# B&R Automation Studio project DemoCNC
Automation Studio 6.7.0.187; technology packages: mappCockpit 6.7.0, mappMotion 6.7.2, mappView 6.7.0, OpcUaCs 6.0.0

## Configuration Config1

CPU X20CP1684, AutomationRuntime 6.7.6, Build 11.3.0, Vc 6.0.0

### Task classes (Cpu.sw)
```
Cyclic#1 (cycle 2000 us, tolerance 0 us):
  Main <- Cnc.Main.prg
  AxisManual <- Motion.AxisManual.prg
  Handwheel <- Motion.Handwheel.prg
  RingBuffer <- Motion.RingBuffer.prg
  Dispenser <- Heads.Dispenser.prg
  Laser <- Heads.Laser.prg
  OpMode <- Cnc.OpMode.prg
Cyclic#4:
  PrgShare <- Cnc.PrgShare.prg
DataObjects: McAcpSys
NcDataObjects: McDriveLog
Binaries: udbdef, ArSvcReg, FWRules, McProfGen, McAcpSim, mvLoader, McAcpDrv, TCData, iomap, Config_4, asfw, Config_3, Settings, Role, Config_6, Config_2, mCoWebSc, User, UaCsConfig, BRRole, Config_5, Config_1, asnxdb1, arconfig, ashwac, ashwd, sysconf
Libraries: runtime, AsZip, FileIO, McBase, MpBase, McAxGroup, McAcpAx, McAxis, McPathGen, MpAxis, McProgInt, McPureVAx, MpCnc, CoTrace, standard, ArSsl, powerlnk, AsIecCon, UaCoal, sys_lib, astime, UaCoalPrv, AsEPL
```

### Hardware
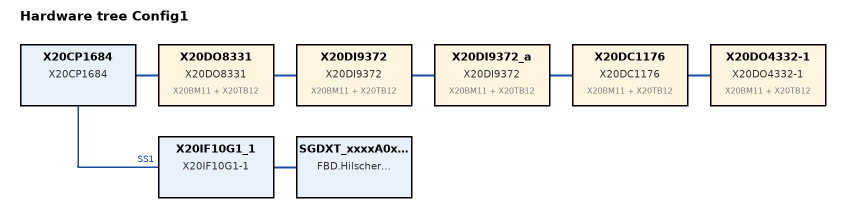
```
SGDXT_xxxxA0x_CoE_Drive_V5_1 : FBD.Hilscher.ECATGenSlaveDTM.SGDXT-xxxxA0x CoE Drive V5.1 v5.1 (OrderNumber=SGDXT-xxxxA0x CoE Drive V5.1)  [ECAT1 -> X20IF10G1_1.IF1]
  DtmId = 5cc0e974-dd08-4d3b-8861-9af8db60d9c1
  ChannelBlocks_556a5014-3061-476e-952f-13eb48db60da  // 2nd_Receive_PDO_mapping_ChA   [OUT, 6 Byte(s)]
  ChannelBlocks_c08b9fef-1a5d-4400-99d8-8c6c7c6492c0  // 2nd_Receive_PDO_mapping_ChB   [OUT, 6 Byte(s)]
  ChannelBlocks_bb719693-a827-4383-9817-184275cbd3ab  // 2nd_Receive_PDO_mapping_ChC   [OUT, 6 Byte(s)]
  ChannelBlocks_bb52f712-f110-4765-9ae9-fe54bf8f2216  // 2nd_Transmit_PDO_mapping_ChA   [IN, 6 Byte(s)]
  ChannelBlocks_06cbf0f9-47c2-45b5-ab43-e0b9d19c4fe2  // 2nd_Transmit_PDO_mapping_ChB   [IN, 6 Byte(s)]
  ChannelBlocks_3a11469b-f58f-4501-9f2d-befe904e9021  // 2nd_Transmit_PDO_mapping_ChC   [IN, 6 Byte(s)]
X20BM11 : X20BM11 v1.1.0.0  [X2X1 -> X20BM11_a.X2X2]
X20BM11_a : X20BM11 v1.1.0.0  [X2X1 -> X20CP1684.IF6]
X20BM11_b : X20BM11 v1.1.0.0  [X2X1 -> X20BM11.X2X2]
X20BM11_c : X20BM11 v1.1.0.0  [X2X1 -> X20BM11_b.X2X2]
X20BM11_d : X20BM11 v1.1.0.0  [X2X1 -> X20BM11_c.X2X2]
X20CP1684 : X20CP1684 v1.9.0.0
  Connector IF2:
    ActivateDevice = 1
    Mode = Manual
    InternetAddress = 192.0.2.10
    SubnetMask = 255.255.255.0
  ConfigurationID = first_Config1
  TimerDeviceType = EPLX2X
  TimerDevice = X20CP1684.IF6
  TaskClassIdleTime = 2000
  Cyclic1Duration = 2000
  Cyclic1Tolerance = 0
  FileDevice1
  FileDeviceName1 = USER
  FileDevicePath1 = USER_PATH
  ActivateWebServer = 1
  ActivateSdm = 1
  Authentication = 0
X20DC1176 : X20DC1176 v1.4.2.0  [SS1 -> X20TB12_c.SS; SL -> X20BM11_c.SL1]
  Supervision = off
  CounterStd01 = 32Bit
  ABRInputs = on
  BrokenWireConfig = off
X20DI9372 : X20DI9372 v1.6.1.0  [SS1 -> X20TB12.SS; SL -> X20BM11.SL1]
  Supervision = off
X20DI9372_a : X20DI9372 v1.6.1.0  [SS1 -> X20TB12_b.SS; SL -> X20BM11_b.SL1]
  Supervision = off
X20DO4332-1 : X20DO4332-1 v1.7.1.0  [SS1 -> X20TB12_d.SS; SL -> X20BM11_d.SL1]
  Supervision = off
X20DO8331 : X20DO8331 v1.2.2.0  [SS1 -> X20TB12_a.SS; SL -> X20BM11_a.SL1]
  Supervision = off
X20IF10G1_1 : X20IF10G1-1 v1.0.2.0  [SS -> X20CP1684.SS1]
  Connector IF1:
    DtmRef = FBDIF.Hilscher.ECATMasterDTM.NETX 100 RE/ECM
    DtmId = 1a6e2b8c-b0d3-41a0-9abf-558976bc5f68
  ConfigFile = X20IF10G1_1.dtm
  ConfigModule = asnxdb1
  CycleTime = 2000
  Synchron = on
X20TB12 : X20TB12 v1.0.0.0
X20TB12_a : X20TB12 v1.0.0.0
X20TB12_b : X20TB12 v1.0.0.0
X20TB12_c : X20TB12 v1.0.0.0
X20TB12_d : X20TB12 v1.0.0.0
```

### BRRole.brrole - X20CP1684/AccessAndSecurity/UserRoleSystem/BRRole.brrole
```
Element BR_Anonymous (Type=BRRole)
Element BR_Engineer (Type=BRRole)
Element BR_Observer (Type=BRRole)
Element BR_SafetyAdmin (Type=BRRole)
Element BR_SecurityAdmin (Type=BRRole)
```

### IoMap.iom - X20CP1684/IoMap.iom
```iecst
VAR_CONFIG
	::gDS402_X.ControlWord AT %QW."SGDXT_xxxxA0x_CoE_Drive_V5_1".2nd_Receive_PDO_mapping_ChA_Control_word;
	::gDS402_X.TargetPosition AT %QD."SGDXT_xxxxA0x_CoE_Drive_V5_1".2nd_Receive_PDO_mapping_ChA_Target_position;
	::gDS402_Y.ControlWord AT %QW."SGDXT_xxxxA0x_CoE_Drive_V5_1".2nd_Receive_PDO_mapping_ChB_Control_word;
	::gDS402_Y.TargetPosition AT %QD."SGDXT_xxxxA0x_CoE_Drive_V5_1".2nd_Receive_PDO_mapping_ChB_Target_position;
	::gDS402_Z.ControlWord AT %QW."SGDXT_xxxxA0x_CoE_Drive_V5_1".2nd_Receive_PDO_mapping_ChC_Control_word;
	::gDS402_Z.TargetPosition AT %QD."SGDXT_xxxxA0x_CoE_Drive_V5_1".2nd_Receive_PDO_mapping_ChC_Target_position;
	::gDS402_X.StatusWord AT %IW."SGDXT_xxxxA0x_CoE_Drive_V5_1".2nd_Transmit_PDO_mapping_ChA_Status_word;
	::gDS402_X.ActualPosition AT %ID."SGDXT_xxxxA0x_CoE_Drive_V5_1".2nd_Transmit_PDO_mapping_ChA_Position_actual_value;
	::gDS402_Y.StatusWord AT %IW."SGDXT_xxxxA0x_CoE_Drive_V5_1".2nd_Transmit_PDO_mapping_ChB_Status_word;
	::gDS402_Y.ActualPosition AT %ID."SGDXT_xxxxA0x_CoE_Drive_V5_1".2nd_Transmit_PDO_mapping_ChB_Position_actual_value;
	::gDS402_Z.StatusWord AT %IW."SGDXT_xxxxA0x_CoE_Drive_V5_1".2nd_Transmit_PDO_mapping_ChC_Status_word;
	::gDS402_Z.ActualPosition AT %ID."SGDXT_xxxxA0x_CoE_Drive_V5_1".2nd_Transmit_PDO_mapping_ChC_Position_actual_value;
	::gDS402_X.DigitalInputs.NegativeLimitSwitch AT %IX."X20DI9372".DigitalInput01;
	::gDS402_X.DigitalInputs.HomingSwitch AT %IX."X20DI9372".DigitalInput02;
	::gDS402_X.DigitalInputs.PositiveLimitSwitch AT %IX."X20DI9372".DigitalInput03;
	::gDS402_Y.DigitalInputs.NegativeLimitSwitch AT %IX."X20DI9372".DigitalInput04;
	::gDS402_Y.DigitalInputs.HomingSwitch AT %IX."X20DI9372".DigitalInput05;
	::gDS402_Y.DigitalInputs.PositiveLimitSwitch AT %IX."X20DI9372".DigitalInput06;
	::gDS402_Z.DigitalInputs.NegativeLimitSwitch AT %IX."X20DI9372".DigitalInput07;
	::gDS402_Z.DigitalInputs.HomingSwitch AT %IX."X20DI9372".DigitalInput08;
	::gDS402_Z.DigitalInputs.PositiveLimitSwitch AT %IX."X20DI9372".DigitalInput09;
	::DO_Dispenser_Start AT %QX."X20DO8331".DigitalOutput01;
	::DO_Laser_Power AT %QX."X20DO8331".DigitalOutput02;
	::PWM_Laser_Duty AT %QW."X20DO4332-1".PwmOutput01;
	::PWM_Laser_Period AT %QW."X20DO4332-1".PwmPeriode;
	::Handwheel:counterValue AT %ID."X20DC1176".Encoder01;
	::Handwheel:counterReset AT %QX."X20DC1176".Encoder01Reset;
	::DI_MPG_AxisX AT %IX."X20DI9372_a".DigitalInput01;
	::DI_MPG_AxisY AT %IX."X20DI9372_a".DigitalInput02;
	::DI_MPG_AxisZ AT %IX."X20DI9372_a".DigitalInput03;
	::DI_MPG_X1 AT %IX."X20DI9372_a".DigitalInput05;
	::DI_MPG_X10 AT %IX."X20DI9372_a".DigitalInput06;
	::DI_MPG_X100 AT %IX."X20DI9372_a".DigitalInput07;
	::DI_MPG_Jog_EMS1 AT %IX."X20DI9372_a".DigitalInput08;
END_VAR
```

- Physical/Config1/X20CP1684/PvMap.vvm: same as Physical/Config1/X20CP1684/Cpu.per
### Config_1.axesgroup - X20CP1684/mappMotion/3AxesCNCXYZ/Config_1.axesgroup
```
Element gCncXYZ (Type=axesgroup)
  Type = PathGenAxesGroup
    PhysicalAxes:
      JointAxes:
        JointAxis[1]:
          Name = QX
          AxisRef = gAxis_X
        JointAxis[2]:
          Name = QY
          AxisRef = gAxis_Y
        JointAxis[3]:
          Name = QZ
          AxisRef = gAxis_Z
    MechanicalSystem:
      MechSysRef = MechSys_3AxCNCXYZ
    AxesGroupFeatures:
      FeatureRef[1] = Feature_Programs
      FeatureRef[2] = Feature_Jogging
      FeatureRef[3] = Feature_MFunctions
      FeatureRef[4] = Feature_HomingOrder
      FeatureRef[5] = Feature_PrgSimAndRestart
```

### Config_2.axis - X20CP1684/mappMotion/3AxesCNCXYZ/Config_2.axis
```
Element gAxis_X (Type=axis)
  BaseType = LinearBounded
    MeasurementResolution = 0.001
    CountDirection = Inverse
  MovementLimits:
    Position:
      LowerLimit = -5
      UpperLimit = 450
    Velocity:
      Velocity = 200
    Acceleration:
      Acceleration = 500.0
    Deceleration:
      Deceleration = 500.0
Element gAxis_Y (Type=axis)
  BaseType = LinearBounded
    MeasurementResolution = 0.001
    CountDirection = Inverse
  MovementLimits:
    Position:
      LowerLimit = -5
      UpperLimit = 430
    Velocity:
      Velocity = 200
    Acceleration:
      Acceleration = 500.0
    Deceleration:
      Deceleration = 500.0
Element gAxis_Z (Type=axis)
  BaseType = LinearBounded
    MeasurementResolution = 0.001
  MovementLimits:
    Position:
      LowerLimit = -5
      UpperLimit = 145
    Velocity:
      Velocity = 200
    Acceleration:
      Acceleration = 500.0
    Deceleration:
      Deceleration = 500.0
```

### Config_3.mechanicalsystem - X20CP1684/mappMotion/3AxesCNCXYZ/Config_3.mechanicalsystem
```
Element MechSys_3AxCNCXYZ (Type=mechanicalsystem)
  Type = 3AxesCNC
    Subtype:
      JointAxesPositionLimits:
        JointAxis[1]
        JointAxis[2]
        JointAxis[3]
```

### Config_4.axesgroupfeature - X20CP1684/mappMotion/3AxesCNCXYZ/Config_4.axesgroupfeature
```
Element Feature_Programs (Type=axesgroupfeature)
  Type = Program
    ModalDataBehaviour = UseAxesGroupSettings
    InitialSettings:
      InterpolationTypes = LinearRapid
      PositionCoordinates = Absolute
      CircleCoordinates = Relative
      JACS_ACSProgramming = JACS
      ContourConnection = Inactive
      AccuracyHoldDelays = None
      ProgrammingUnits = UseAxesGroupSettings
      Feedrates:
        FeedPath = Standard
        FeedCharacteristic = StandardCharacteristic
        FeedType = Feedrate
        FeedReduction = Inactive
        FeedrateValue = 0.0
        InverseFeedrateValue = 0.0
        FeedratePerRevValue = 0.0
    ProgramElements:
      PVs:
        PV[1]:
          PvName = ::C_LaserPower
          Advanced:
            Alias = LaserPower
            Synchronization = Path
        PV[2]:
          PvName = ::C_TP1_1
          Advanced:
            Alias = TP1_1
        PV[3]:
          PvName = ::C_TP1_2
          Advanced:
            Alias = TP1_2
        PV[4]:
          PvName = ::C_TP1_3
          Advanced:
            Alias = TP1_3
        PV[5]:
          PvName = ::C_TP2_1
          Advanced:
            Alias = TP2_1
        PV[6]:
          PvName = ::C_TP2_2
          Advanced:
            Alias = TP2_2
        PV[7]:
          PvName = ::C_TP2_3
          Advanced:
            Alias = TP2_3
        PV[8]:
          PvName = ::C_TP3_1
          Advanced:
            Alias = TP3_1
        PV[9]:
          PvName = ::C_TP3_2
          Advanced:
            Alias = TP3_2
        PV[10]:
          PvName = ::C_TP3_3
          Advanced:
            Alias = TP3_3
        PV[11]:
          PvName = ::C_TP4_1
          Advanced:
            Alias = TP4_1
        PV[12]:
          PvName = ::C_TP4_2
          Advanced:
            Alias = TP4_2
        PV[13]:
          PvName = ::C_TP4_3
          Advanced:
            Alias = TP4_3
    DefaultLanguage = BRGCode
    Location = Default
      FileDevice = CNC_PrgDir
Element Feature_Jogging (Type=axesgroupfeature)
  Type = Jogging
```

### Config_5.purevaxcfg - X20CP1684/mappMotion/3AxesCNCXYZ/Config_5.purevaxcfg
```
Element PureVAxCfg_X (Type=purevaxcfg)
  PureVAxis:
    AxisReference = gAxis_X
    Homing:
      Mode = SwitchGate
        SwitchEdge = Negative
        StartDirection = Negative
    GeneralPurposeAxisInterface = DS402CSP
      MechanicalElements:
        RotaryToLinearTransformation:
          ReferenceDistance = 10
      EncoderSettings:
        IncrementsPerRevolution = 1048576
      PositionActualValue:
        Source = Variable
          PVMapping = ::gDS402_X.ActualPosition
      DigitalInputs:
        HomingSwitch:
          Source = InputPV
            PVmapping = ::gDS402_X.DigitalInputs.HomingSwitch
        PositiveLimitSwitch:
          Source = InputPV
            PVmapping = ::gDS402_X.DigitalInputs.PositiveLimitSwitch
          Level = Low
        NegativeLimitSwitch:
          Source = InputPV
            PVmapping = ::gDS402_X.DigitalInputs.NegativeLimitSwitch
          Level = Low
      StatusInputs:
        StatusWord:
          Source = InputPV
            PVmapping = ::gDS402_X.StatusWord
        ErrorCode:
          Source = InputPV
            PVmapping = ::gDS402_X.ErrorCode
      ControlOutputs:
        ControlWord:
          Destination:
            PVMapping = ::gDS402_X.ControlWord
        TargetPosition:
          Destination:
            PVmapping = ::gDS402_X.TargetPosition
Element PureVAxCfg_Y (Type=purevaxcfg)
  PureVAxis:
    AxisReference = gAxis_Y
    Homing:
      Mode = SwitchGate
        Position = 0
        SwitchEdge = Negative
        StartDirection = Negative
    GeneralPurposeAxisInterface = DS402CSP
      MechanicalElements:
        RotaryToLinearTransformation:
          ReferenceDistance = 10
      EncoderSettings:
        IncrementsPerRevolution = 1048576
      PositionActualValue:
        Source = Variable
          PVMapping = ::gDS402_Y.ActualPosition
      DigitalInputs:
        HomingSwitch:
          Source = InputPV
            PVmapping = ::gDS402_Y.DigitalInputs.HomingSwitch
        PositiveLimitSwitch:
          Source = InputPV
            PVmapping = ::gDS402_Y.DigitalInputs.PositiveLimitSwitch
          Level = Low
        NegativeLimitSwitch:
          Source = InputPV
            PVmapping = ::gDS402_Y.DigitalInputs.NegativeLimitSwitch
          Level = Low
      StatusInputs:
        StatusWord:
          Source = InputPV
            PVmapping = ::gDS402_Y.StatusWord
        ErrorCode:
          Source = InputPV
            PVmapping = ::gDS402_Y.ErrorCode
      ControlOutputs:
        ControlWord:
          Destination:
            PVMapping = ::gDS402_Y.ControlWord
        TargetPosition:
          Destination:
            PVmapping = ::gDS402_Y.TargetPosition
Element PureVAxCfg_Z (Type=purevaxcfg)
  PureVAxis:
    AxisReference = gAxis_Z
    Homing:
      Mode = SwitchGate
        SwitchEdge = Negative
        StartDirection = Negative
    GeneralPurposeAxisInterface = DS402CSP
      MechanicalElements:
        RotaryToLinearTransformation:
          ReferenceDistance = 10
      EncoderSettings:
        IncrementsPerRevolution = 1048576
      PositionActualValue:
        Source = Variable
          PVMapping = ::gDS402_Z.ActualPosition
      DigitalInputs:
        HomingSwitch:
          Source = InputPV
            PVmapping = ::gDS402_Z.DigitalInputs.HomingSwitch
        PositiveLimitSwitch:
          Source = InputPV
            PVmapping = ::gDS402_Z.DigitalInputs.PositiveLimitSwitch
          Level = Low
        NegativeLimitSwitch:
          Source = InputPV
            PVmapping = ::gDS402_Z.DigitalInputs.NegativeLimitSwitch
          Level = Low
      StatusInputs:
        StatusWord:
          Source = InputPV
            PVmapping = ::gDS402_Z.StatusWord
        ErrorCode:
          Source = InputPV
            PVmapping = ::gDS402_Z.ErrorCode
      ControlOutputs:
        ControlWord:
          Destination:
            PVMapping = ::gDS402_Z.ControlWord
        TargetPosition:
          Destination:
            PVmapping = ::gDS402_Z.TargetPosition
```

### Config_6.axesgroupfeature - X20CP1684/mappMotion/3AxesCNCXYZ/Config_6.axesgroupfeature
```
Element Feature_MFunctions (Type=axesgroupfeature)
  Type = MFunctions
    MFunction[1]:
      IndexType = Range
        IndexFrom = 40
        IndexTo = 49
      Blocking = Disabled
    MFunction[2]:
      IndexType = Range
        IndexFrom = 50
        IndexTo = 59
    MFunction[3]:
      IndexType = Range
        IndexFrom = 60
        IndexTo = 69
      Blocking = Disabled
```

### Config_7.axesgroupfeature - X20CP1684/mappMotion/3AxesCNCXYZ/Config_7.axesgroupfeature
```
Element Feature_HomingOrder (Type=axesgroupfeature)
  Type = HomingOrder
    TogetherGroup[1]:
      AxisRef[1] = gAxis_Z
    TogetherGroup[2]:
      AxisRef[1] = gAxis_X
      AxisRef[2] = gAxis_Y
```

### Config_8.axesgroupfeature - X20CP1684/mappMotion/3AxesCNCXYZ/Config_8.axesgroupfeature
```
Element Feature_PrgSimAndRestart (Type=axesgroupfeature)
  Type = SimulationRestart
    ConditionalStop = NotUsed
    AdvancedParameters = NotUsed
```

## Logical view

Binary libraries used (declarations not repeated): operator, runtime, AsIecCon, astime, AsZip, FileIO, McBase 6.7.2, MpBase 6.5.0, McAxGroup 6.7.2, McAcpAx 6.7.2, McAxis 6.7.2, McPathGen 6.7.2, MpAxis 6.7.2, McProgInt 6.7.2, McPureVAx 6.7.2, MpCnc 6.7.2, CoTrace 6.7.0, standard

### Global.typ - Global data types
```iecst
TYPE
	Equip_Type : 	STRUCT
		Input : EquipInput_Type;
		Output : EquipOutput_Type;
	END_STRUCT;
	EquipInput_Type : 	STRUCT
		Command : EquipInputCommand_Type;
		CncCommand : E_CNC_ACTION;
		Parameter : EquipInputParameter_Type;
	END_STRUCT;
	EquipOutput_Type : 	STRUCT
		State : EquipOutputState_Type;
		Status : EquipOutputStatus_Type;
	END_STRUCT;
	EquipInputCommand_Type : 	STRUCT
		ManualMove : BOOL; (*move to Parameter.ManualPositon (Z retracts to 0 first) - manual mode, homed*)
		AlarmClearAll : BOOL;
		ManualMode : BOOL; (*TRUE = manual mode (jog, position move, manual discharge). Ignored while the CNC is busy*)
	END_STRUCT;
	EquipInputParameter_Type : 	STRUCT
		sProgramName : STRING[80];
		DryRun : BOOL;
		SystemSpeed : REAL;
		Feedrate : REAL;
		ManualSlowMove : BOOL;
		ManualPositon : ARRAY[0..2]OF REAL;
		sBlock : STRING[260]; (*single NC block for E_ACT_MOVE_BLOCK (MDI), e.g. 'G90 G01 X10 Y20 F1000'*)
		sInitProgram : STRING[80]; (*init program run before every program START (not MDI) as an init subroutine of the program (MoveProgramOptions.InitProgram), e.g. a G92 or a move to a teach position. Empty = none*)
	END_STRUCT;
	EquipOutputState_Type : 	STRUCT
		Initialized : BOOL;
		Stop : BOOL;
		Move : BOOL;
		Complete : BOOL;
	END_STRUCT;
	EquipOutputStatus_Type : 	STRUCT
		CurrentAction : E_CNC_ACTION;
		Mode : BOOL;
		ManualMove : BOOL;
		MoveComplete : BOOL;
		WorkPanelName : STRING[255];
		PowerOn : BOOL; (*CNC axes powered*)
		IsHomed : BOOL; (*CNC axes homed - FALSE after every power-up until HOME / INIT*)
		ProgramActive : BOOL; (*CNC program executing (also while interrupted)*)
		ProgramInterrupted : BOOL; (*CNC program interrupted by HALT*)
		Error : BOOL; (*MpCnc3Axis error*)
		StatusID : DINT; (*MpCnc3Axis StatusID*)
		Rejected : E_CNC_ACTION; (*last mailbox command discarded because its preconditions were not met, IDLE after an accepted command*)
		EmergencyStop : BOOL; (*E-stop latched - release the button, then RESET*)
	END_STRUCT;
	E_CNC_ACTION :
		(
		E_ACT_IDLE := 0,
		E_ACT_INIT := 1,
		E_ACT_START := 2,
		E_ACT_HALT := 3,
		E_ACT_STOP := 4,
		E_ACT_RESET := 5,
		E_ACT_CONTINUE := 6,
		E_ACT_LOADPROGRAM := 7,
		E_ACT_HOME := 8,
		E_ACT_ABORT := 10, (*leave the running command without an action (Main), refused while idle*)
		E_ACT_POWER_OFF := 13, (*servo off*)
		E_ACT_MOVE_BLOCK := 14, (*execute Parameter.sBlock (MDI)*)
		E_ACT_START_AT_LINE := 15, (*START from the file line gCncRun.Input.StartLine*)
		E_ACT_MEASURE_Z := 16 (*Z reference measurement with the touch sensor (gZRef) - manual mode, homed*)
		);
END_TYPE

(*Dispenser*)

TYPE
	Dispenser_Type : 	STRUCT
		Input : DispenserInput_Type;
		Output : DispenserOutput_Type;
	END_STRUCT;
	DispenserInput_Type : 	STRUCT
		Command : DispenserInputCommand_Type;
		Parameter : DispenserInputParameter_Type;
	END_STRUCT;
	DispenserOutput_Type : 	STRUCT
		State : DispenserOutputState_Type;
	END_STRUCT;
	DispenserInputCommand_Type : 	STRUCT
		Discharge : BOOL; (*auto : M41 on / M42 off, driven by Main*)
		Manual : BOOL; (*manual on/off*)
	END_STRUCT;
	DispenserInputParameter_Type : 	STRUCT
		DischargeDelay : BOOL; (*M44 on / M45 off - flag for the program, no output function on this machine*)
	END_STRUCT;
	DispenserOutputState_Type : 	STRUCT
		Discharge : BOOL; (*TRUE while the dispenser discharges (DO_Dispenser_Start)*)
	END_STRUCT;
END_TYPE

(*Laser*)

TYPE
	Laser_Type : 	STRUCT
		Input : LaserInput_Type;
		Output : LaserOutput_Type;
	END_STRUCT;
	LaserInput_Type : 	STRUCT
		Command : LaserInputCommand_Type;
		Parameter : LaserInputParameter_Type;
	END_STRUCT;
	LaserOutput_Type : 	STRUCT
		State : LaserOutputState_Type;
	END_STRUCT;
	LaserInputCommand_Type : 	STRUCT
		Emission : BOOL; (*auto : M61 on / M62 off, driven by Main*)
		Manual : BOOL; (*manual on/off*)
	END_STRUCT;
	LaserInputParameter_Type : 	STRUCT (*written by the HMI (gLaser is not RETAIN, the Laser Init sets the start values)*)
		Power : REAL; (*auto power [%] while the program sets no LaserPower (C_LaserPower < 0)*)
		ManualPower : REAL; (*manual test power [%]*)
		DutyMin : REAL; (*PWM duty for a power just above 0 % [%] - lasing threshold of the driver*)
		DutyMax : REAL; (*PWM duty for 100 % power [%]*)
		PwmPeriod : UINT; (*PWM period [us], 1000..65535 (1000 = 1 kHz, the X20DO4332-1 maximum)*)
		SpeedScale : BOOL; (*corner compensation : power x actual / programmed path velocity*)
		MinSpeedRatio : REAL; (*lower limit of that velocity ratio [%]*)
	END_STRUCT;
	LaserOutputState_Type : 	STRUCT
		Emission : BOOL; (*TRUE while the laser emits (DO_Laser_On : on and power > 0)*)
		Power : REAL; (*power output now [%], after corner compensation, 0 while off*)
		Duty : REAL; (*PWM duty output now [%]*)
	END_STRUCT;
END_TYPE

(*Axis*)

TYPE
	AXIS_COMMAND :
		(
		Axis_IDLE := 0,
		Axis_MOVE_ABSOLUTE := 1,
		Axis_STOP := 2,
		Axis_HALT := 3,
		Axis_JOG_NEGATIVE := 4,
		Axis_JOG_POSITIVE := 5,
		Axis_RESET := 6,
		Axis_MOVE_ADDITIVE := 7,
		Axis_HOME := 8,
		Axis_POWER := 9,
		Axis_MOVE_VELOCITY := 10
		);
	AxesInterface_Type : 	STRUCT
		Input : AxisInput_Type;
		Output : AxisOutput_Type;
	END_STRUCT;
	AxisInput_Type : 	STRUCT
		Parameter : AxisParameter_Type;
		Command : AxisCommand_Type;
	END_STRUCT;
	AxisOutput_Type : 	STRUCT
		State : AxisState_Type;
	END_STRUCT;
	AxisCommand_Type : 	STRUCT
		JogNegative : BOOL;
		JogPositive : BOOL;
		Reset : BOOL;
		Command : AXIS_COMMAND;
	END_STRUCT;
	AxisParameter_Type : 	STRUCT
		Speed : REAL;
		Position : REAL;
		Distance : REAL;
		JogSpeed : REAL;
		SoftwareLimitsPos : DINT;
		SoftwareLimitsNeg : DINT;
		Power : BOOL; (*target of Axis_POWER : TRUE = on, FALSE = off*)
	END_STRUCT;
	AxisState_Type : 	STRUCT
		Enable : BOOL;
		Home : BOOL;
		JogNegative : BOOL;
		JogPositive : BOOL;
		Error : BOOL;
		ErrorID : UDINT;
		Status : SINT; (*0: Not Init , 1 : Idle or OK , 2 : Run, 3 : Error *)
		Command : AXIS_COMMAND;
		Position : LREAL;
		Speed : LREAL;
	END_STRUCT;
END_TYPE

(*Drive diagnosis - read-only copies for the HMI, not RETAIN (gAxis is RETAIN and keeps its structure). Written by AxisManual*)

TYPE
	DriveDiag_Type : 	STRUCT
		Valid : BOOL; (*the values below are up to date (MC_ReadAxisInfo.Valid) - FALSE = do not judge them*)
		CommReady : BOOL; (*drive has a network connection (MC_ReadAxisInfo.CommunicationReady) - follows the 'Module ok' status input of the axis config (Config_5), not used yet*)
		ReadyForPowerOn : BOOL; (*drive can be switched on (MC_ReadAxisInfo.ReadyForPowerOn)*)
		Warning : BOOL; (*a warning is active on the drive (MC_ReadAxisInfo.AxisWarning, DS402 status word bit 7)*)
		WarningAlarm : BOOL; (*warning-level alarm for the HMI (alarms.json exType 1) : Warning while Valid and CommReady for 0.5 s, held 2 s after it clears (one alarm per event, no flicker). Display only - the PLC does not react to it*)
	END_STRUCT;
END_TYPE

(*Position move result*)

TYPE
	ManualMoveResult_Type : 	STRUCT (*result of gEquipment.Input.Command.ManualMove, written by AxisManual - its own non-RETAIN global so the RETAIN gEquipment keeps its layout*)
		Result : USINT; (*result of request number Count : 0 none since power-up, 1 running, 2 arrived (every step of the sequence done), 3 refused (dropped, nothing moved), 4 ended before the target (Reason)*)
		Reason : USINT; (*why refused / ended, 0 none : 1 E-stop, 2 auto mode, 3 handwheel selected, 4 CNC command running, 5 axes moving, 6 not homed, 7 servo off, 8 axis error, 9 axis HALT / STOP, 10 an axis move of the sequence was aborted or failed (the sequence went on)*)
		Count : UINT; (*+1 for every ManualMove request the PLC takes (accepted or refused) : a new result also when it equals the last one*)
	END_STRUCT;
END_TYPE

(*Z reference measurement - touch sensor DI_ZRef_Sensor (not wired yet), cycle in Main Action_ZRef.st (CncCommand E_ACT_MEASURE_Z)*)

TYPE
	ZRef_Type : 	STRUCT
		Input : ZRefInput_Type;
		Output : ZRefOutput_Type;
	END_STRUCT;
	ZRefInput_Type : 	STRUCT (*written by the HMI, kept over power off (gZRef is RETAIN) - machine coordinates [mm], Z+ down (0 = top). All 0 = not set : the command is refused*)
		SensorX : LREAL; (*X of the sensor*)
		SensorY : LREAL; (*Y of the sensor*)
		StartZ : LREAL; (*Z above the sensor where the slow search starts*)
		MaxZ : LREAL; (*deepest Z of the search : no signal down to here = failed (at most 50 mm below StartZ)*)
		SafeZ : LREAL; (*Z of the moves to and from the sensor (not below StartZ), usually 0*)
		ProbeVel : REAL; (*search velocity [mm/s], 0 = 2, at most 10. The result is read once per cycle : error up to about ProbeVel x 2 cycles (2 ms) + the input filter*)
		Head : USINT; (*head being measured (HMI head number), copied to Output.Head with the result*)
	END_STRUCT;
	ZRefOutput_Type : 	STRUCT
		ParamOk : BOOL; (*Input valid : SafeZ <= StartZ < MaxZ, search <= 50 mm, all inside the software limits, ProbeVel <= 10*)
		Sensor : BOOL; (*DI_ZRef_Sensor now*)
		Busy : BOOL; (*measurement running*)
		Step : USINT; (*diagnosis: 10 Z to SafeZ, 20 X / Y to the sensor, 30 Z to StartZ, 40 search, 50 braking, 60 Z back to SafeZ*)
		Done : BOOL; (*MeasuredZ is the result of the last measurement (cleared when the next one starts)*)
		MeasuredZ : LREAL; (*Z at the sensor signal [mm, machine]*)
		Head : USINT; (*head of MeasuredZ*)
		ErrorId : USINT; (*last measurement: 0 none, 1 Input not valid, 2 sensor already on at StartZ, 3 no signal down to MaxZ, 4 axis move failed or aborted (jog, axis error), 5 left (STOP, ABORT, E-stop, handwheel), 6 a move did not finish in time*)
	END_STRUCT;
END_TYPE

(*Work offsets G54..G57 - program origin in machine coordinates, set as the standard frame SCS1 before a program / MDI run (Main Action_WorkOffset.st)*)

TYPE
	WorkOffset_Type : 	STRUCT
		Input : WorkOffsetInput_Type;
		Output : WorkOffsetOutput_Type;
	END_STRUCT;
	WorkOffsetInput_Type : 	STRUCT
		Command : WorkOffsetInputCommand_Type;
		Parameter : WorkOffsetInputParameter_Type;
	END_STRUCT;
	WorkOffsetInputCommand_Type : 	STRUCT
		Apply : BOOL; (*pulse: take Parameter over (table and Active), cleared by the PLC - refused while a command / program runs*)
	END_STRUCT;
	WorkOffsetInputParameter_Type : 	STRUCT
		Offset : ARRAY[0..3]OF WorkOffsetXYZ_Type; (*0 = G54 .. 3 = G57 : machine position of the program origin [mm]*)
		Active : USINT; (*0..3 = G54..G57 : offset used by every program and MDI run*)
	END_STRUCT;
	WorkOffsetXYZ_Type : 	STRUCT
		X : LREAL;
		Y : LREAL;
		Z : LREAL;
	END_STRUCT;
	WorkOffsetOutput_Type : 	STRUCT
		Offset : ARRAY[0..3]OF WorkOffsetXYZ_Type; (*table in effect (taken over by Apply, kept over power off)*)
		Active : USINT; (*offset in effect, 0 = G54*)
		InUse : BOOL; (*the frame is set before every run : the active offset or the frame set last is not 0*)
		Rejected : BOOL; (*the last Apply was refused : CNC busy, Active > 3 or a value out of range (10000 mm)*)
		Error : BOOL; (*setting the frame failed - that run was not started*)
		ErrorID : DINT; (*ErrorID of MC_BR_SetStandardFrame, 0 = none*)
	END_STRUCT;
END_TYPE

(*Head (tool) offsets - offset of the mounted head from the reference head tip, set as the standard frame SCS2 before a program / MDI run (Main Action_HeadOffset.st)*)

TYPE
	HeadOffset_Type : 	STRUCT
		Input : HeadOffsetInput_Type;
		Output : HeadOffsetOutput_Type;
	END_STRUCT;
	HeadOffsetInput_Type : 	STRUCT
		Command : HeadOffsetInputCommand_Type;
		Parameter : HeadOffsetInputParameter_Type;
	END_STRUCT;
	HeadOffsetInputCommand_Type : 	STRUCT
		Apply : BOOL; (*pulse: take Parameter over (table and ActiveHead), cleared by the PLC - refused while a command / program runs*)
	END_STRUCT;
	HeadOffsetInputParameter_Type : 	STRUCT
		Offset : ARRAY[1..4]OF HeadOffsetXYZ_Type; (*head 1..4 (HMI head table H1..H4 = plugin PlcId : 1 dispenser, 2 laser) : from the reference head tip (the point the axis positions refer to) to the working point of that head [mm], machine directions (Z+ down)*)
		ActiveHead : USINT; (*mounted head 1..4 whose offset every program and MDI run uses, 0 = none (no offset)*)
	END_STRUCT;
	HeadOffsetXYZ_Type : 	STRUCT
		X : LREAL;
		Y : LREAL;
		Z : LREAL;
	END_STRUCT;
	HeadOffsetOutput_Type : 	STRUCT
		Offset : ARRAY[1..4]OF HeadOffsetXYZ_Type; (*table in effect (taken over by Apply, kept over power off)*)
		ActiveHead : USINT; (*head in effect, 0 = none*)
		InUse : BOOL; (*the frame is set before every run : the active head's offset or the frame set last is not 0*)
		Rejected : BOOL; (*the last Apply was refused : CNC busy, ActiveHead > 4 or a value out of range (1000 mm)*)
		Error : BOOL; (*setting the frame failed - that run was not started*)
		ErrorID : DINT; (*ErrorID of MC_BR_SetStandardFrame, 0 = none*)
	END_STRUCT;
END_TYPE

(*CNC program run options from the HMI (gCncRun, not RETAIN : everything is off after a power-up)*)

TYPE
	CncRun_Type : 	STRUCT
		Input : CncRunInput_Type;
		Output : CncRunOutput_Type;
	END_STRUCT;
	CncRunInput_Type : 	STRUCT
		SingleStep : BOOL; (*TRUE = single step : the program stops after every block, CONTINUE runs the next one (MpCnc3Axis.SingleStep). Not used for MDI*)
		OptionalStop : BOOL; (*TRUE = the program stops at M01, CONTINUE goes on (MC_BR_OptionalStop)*)
		StartLine : UDINT; (*E_ACT_START_AT_LINE : line of the program file to start at, 1 = first line (as C_CurrentLine). Write it before CncCommand 15*)
		ReposVelocityFactor : REAL; (*E_ACT_START_AT_LINE : AxisVelocityFactor of the automatic repositioning to the start point (mcPRGRP_SINGLE_AXIS_AUTOMATIC), Main Init sets 0.1*)
	END_STRUCT;
	CncRunOutput_Type : 	STRUCT
		SingleStepActive : BOOL; (*single step mode active (MpCnc3Axis.SingleStepActive)*)
		OptionalStopActive : BOOL; (*the program stands at M01 (MC_BR_OptionalStop.Interrupting) - CONTINUE goes on*)
		OptionalStopErrorId : DINT; (*ErrorID of MC_BR_OptionalStop, 0 = none - switch OptionalStop off and on again to retry*)
		InterruptStatus : McPrgInfoInterruptEnum; (*why the program is interrupted (MpCnc3Axis Info.Program.InterruptStatus) - for commissioning*)
		ProgramPhase : McPrgPhaseEnum; (*MpCnc3Axis Info.Program.ProgramPhase : start at line = simulation up to the line, repositioning, waiting for CONTINUE, real run*)
	END_STRUCT;
END_TYPE
```

### Global.var - Global variables
```iecst
(*Drive adapter - motor / drive specific.
  On a motor or drive change only this block, IoMap.iom, the mappMotion axis configs and the DTM change.
  Program logic uses only the mapp axis references gAxis_X/Y/Z and the axes group gCncXYZ.*)
VAR
	gDS402_X : McPureVAxDS402CspAdapterPvType;
	gDS402_Y : McPureVAxDS402CspAdapterPvType;
	gDS402_Z : McPureVAxDS402CspAdapterPvType;
END_VAR
VAR RETAIN
	gEquipment : Equip_Type;
	gAxis : ARRAY[0..2] OF AxesInterface_Type;
END_VAR
VAR
	gDispenser : Dispenser_Type;
	gLaser : Laser_Type;
END_VAR
(*Axis index of gAxis, gDriveDiag and the per-axis FB arrays*)
VAR CONSTANT
	AX_X : USINT := 0;
	AX_Y : USINT := 1;
	AX_Z : USINT := 2;
	AX_LAST : USINT := 2; (*highest axis index : FOR i := 0 TO AX_LAST*)
END_VAR
(*Drive diagnosis for the HMI - read only (AxisManual overwrites it every cycle), not RETAIN, index AX_X/AX_Y/AX_Z as gAxis*)
VAR
	gDriveDiag : ARRAY[0..2] OF DriveDiag_Type;
END_VAR
(*HMI jog heartbeat - not RETAIN*)
VAR
	gJogAlive : UINT := 0; (*the HMI changes it every 0.1 s while it jogs; AxisManual stops the jog when it stands still for 0.5 s*)
END_VAR
(*Position move result for the HMI - not RETAIN (gEquipment is RETAIN and keeps its layout)*)
VAR
	gManualMoveResult : ManualMoveResult_Type; (*result of the last Input.Command.ManualMove request, written by AxisManual*)
END_VAR
(*Heads - one head on the machine (HMI plugin structure). Head number = PlcId of the HMI head plugin*)
VAR CONSTANT
	HEAD_DISPENSER : USINT := 1; (*dispenser : M41 / M42 discharge on / off, M44 / M45 discharge delay flag, Dispenser task*)
	HEAD_LASER : USINT := 2; (*PWM laser : M61 / M62 emission on / off, Laser task*)
END_VAR
(*Heads this PLC program has - not RETAIN, read by the HMI*)
VAR
	gHeadSupport : UDINT := 0; (*bit n = head n (HEAD_ constants) has its M functions and outputs here. Fixed, set by Main every cycle. The HMI does not offer a head without its bit*)
END_VAR
(*Active head - written by the HMI, not RETAIN. Not in gEquipment : a new field would change the RETAIN structure*)
VAR
	gActiveHead : USINT := 0; (*head selected on the HMI (HEAD_ constant, the plugin PlcId). Only its M functions and manual on are taken : an M function of another head stops the program, a manual on of another head is dropped (Main act_HeadCheck). 0 = not known yet (PLC restart until the HMI writes it) : no check*)
	gHeadRefused : USINT := 0; (*head whose M function or manual on was refused last because it is not gActiveHead (HEAD_ constants), 0 = none. Cleared when the next run starts or by RESET*)
END_VAR
(*CNC program run options from the HMI (single step, M01 stop, start at line) - not RETAIN : off after every power-up*)
VAR
	gCncRun : CncRun_Type;
END_VAR
(*Setting Variable*)
VAR RETAIN
	SlowMoveVelocity : DINT := 10;
	SlowMoveLength : DINT := 100;
END_VAR
(*Monitor*)
VAR
	C_CurrentLine : DINT := 0; (*line of the running CNC program, from MpCnc3Axis ProgramMonitor*)
	C_OverallRuntime : LREAL := 0.0; (*execution time of the running CNC program [s], from MpCnc3Axis ProgramMonitor - counts from the start (file load included) and holds after the end*)
	C_MovementRuntime : LREAL := 0.0; (*movement time of the running CNC program [s], from MpCnc3Axis ProgramMonitor - file load not included*)
	Torque_X : REAL := 0.0;
	Torque_Y : REAL := 0.0;
	Torque_Z : REAL := 0.0;
END_VAR
(*CNC program variables - written by the program through an alias of the axes group program feature (Config_4, path synchronous)*)
VAR
	C_LaserPower : REAL := -1.0; (*LaserPower = <%> in the program; < 0 = not set (gLaser.Input.Parameter.Power), reset at program end*)
END_VAR
(*Teach positions 1..4 [mm, machine coordinates] - read by CNC programs as TP1_1 .. TP4_3 (aliases in Config_4, _1 = X, _2 = Y, _3 = Z : a name
  must not contain X/Y/Z/F after its first letter - an address letter inside an expression
  splits the expression, e.g. 'X=2930-DoubleBeadY=40'), e.g. in the init program
  (Input.Parameter.sInitProgram) 'G00 X=TP1_1 Y=TP1_2' to go there, or 'G92 X=TP4_1 Y=TP4_2' (G92 = absolute zero offset : teach position 4 becomes the program origin). The HMI owns the values (Config\TeachPositions.xml, slot = order
  in Config\Machine.xml) and writes them here whenever they differ*)
VAR RETAIN
	C_TP1_1 : LREAL := 0.0;
	C_TP1_2 : LREAL := 0.0;
	C_TP1_3 : LREAL := 0.0;
	C_TP2_1 : LREAL := 0.0;
	C_TP2_2 : LREAL := 0.0;
	C_TP2_3 : LREAL := 0.0;
	C_TP3_1 : LREAL := 0.0;
	C_TP3_2 : LREAL := 0.0;
	C_TP3_3 : LREAL := 0.0;
	C_TP4_1 : LREAL := 0.0;
	C_TP4_2 : LREAL := 0.0;
	C_TP4_3 : LREAL := 0.0;
END_VAR
(*Z reference measurement (CncCommand E_ACT_MEASURE_Z, Main Action_ZRef.st) - RETAIN on its own (sensor position), gEquipment is
  not changed. The HMI writes Input (sensor position, search range) and reads Output (MeasuredZ, Done, ErrorId)*)
VAR RETAIN
	gZRef : ZRef_Type;
END_VAR
(*Work offsets G54..G57 (Main Action_WorkOffset.st) - RETAIN on its own, gEquipment is not changed. The HMI writes Input.Parameter
  (machine position of the program origin per offset, active offset) and sets Input.Command.Apply while the CNC is idle; the values
  in effect are Output.Offset / Output.Active. All 0 (the default) = program coordinates are machine coordinates*)
VAR RETAIN
	gWorkOffset : WorkOffset_Type;
END_VAR
(*Head (tool) offsets (Main Action_HeadOffset.st) - RETAIN on its own, gEquipment is not changed. The HMI writes Input.Parameter
  (offset per head from the reference head tip, mounted head) and sets Input.Command.Apply while the CNC is idle; the values in
  effect are Output.Offset / Output.ActiveHead. ActiveHead 0 or offset 0 (the default) = no shift*)
VAR RETAIN
	gHeadOffset : HeadOffset_Type;
END_VAR
(*I/O - wired signals only. Axis limit/home switches go straight to gDS402_* in IoMap.iom*)
VAR
	DI_Auto : BOOL := FALSE;
	DI_MPG_AxisX : BOOL := FALSE;
	DI_MPG_AxisY : BOOL := FALSE;
	DI_MPG_AxisZ : BOOL := FALSE;
	DI_MPG_X1 : BOOL := FALSE;
	DI_MPG_X10 : BOOL := FALSE;
	DI_MPG_X100 : BOOL := FALSE;
	DI_MPG_Jog_EMS1 : BOOL := FALSE;
	DI_MPG_Jog_Enable : BOOL := FALSE;
	DO_Dispenser_Start : BOOL := FALSE;
	DO_Laser_Power : BOOL := FALSE; (*X20DO8331 DO02 - on/off laser output, not used by the PWM laser : held FALSE*)
	PWM_Laser_Duty : INT := 0; (*X20DO4332-1 PwmOutput01 : 0..32767 = 0..100 % of the period (power and on/off)*)
	PWM_Laser_Period : UINT := 1000; (*X20DO4332-1 PwmPeriode [us]*)
END_VAR
(*Z reference touch sensor - NOT wired yet : no channel in Hardware.hw / IoMap.iom. Map it in IoMap.iom once the sensor is wired
  (TRUE = touched : an NC sensor needs a NOT where Main reads it). Until then it stays FALSE and a measurement ends at MaxZ (ErrorId 3)*)
VAR
	DI_ZRef_Sensor : BOOL := FALSE;
END_VAR
(*Laser emitting (on and power > 0) - not wired, for the HMI (head lamp, PLC presence)*)
VAR
	DO_Laser_On : BOOL := FALSE;
END_VAR
```


### Package Logical/Cnc - CNC sequence, operating mode, program folder

### Program Logical/Cnc/Main (IEC) - CNC sequencer (MpCnc3Axis)

#### Init.st - Init code
```iecst
PROGRAM _INIT

	gEquipment.Input.CncCommand := E_ACT_IDLE;

	gEquipment.Output.State.Initialized := FALSE;
	gEquipment.Input.Parameter.SystemSpeed := 200; (* [mm/s] position move speed - axis velocity limit is 200 (mappMotion Config_2) *)
	gEquipment.Input.Parameter.Feedrate := 100;

	(* mapp Motion CNC : static references *)
	fbCnc.MpLink := ADR(gCncXYZ);
	fbCnc.Parameters := ADR(CncParameters);
	fbCnc.Enable := TRUE;
	fbCnc.Override := 100.0;
	fbCnc.RapidOverride := 100.0;
	fbCnc.FeedrateOverride := 100.0;

	(* Jog path limits : adjust to machine limits *)
	CncParameters.Jog.PathLimits.Velocity := 1000.0;			(* [mm/s] *)
	CncParameters.Jog.PathLimits.Acceleration := 5000.0;		(* [mm/s^2] *)
	CncParameters.Jog.PathLimits.Deceleration := 5000.0;		(* [mm/s^2] *)

	(* M-Functions : async (AxesGroup M-function feature, ranges 40..49 / 60..69 non-blocking), M50 / M51 blocking (50..59, no function) *)
	fbMFunction[0].MFunction := 41;
	fbMFunction[1].MFunction := 42;
	fbMFunction[2].MFunction := 44;
	fbMFunction[3].MFunction := 45;
	fbMFunction[4].MFunction := 61;
	fbMFunction[5].MFunction := 62;
	fbMFunction[6].MFunction := 50;
	fbMFunction[7].MFunction := 51;
	FOR i := 0 TO 7 DO
		fbMFunction[i].AxesGroup := ADR(gCncXYZ);
		fbMFunction[i].Enable := TRUE;
	END_FOR
	(* M52..M59 : no function here too, act_MSpare lets the path go on (blocking codes of the range would wait for ever) *)
	FOR i := 0 TO 7 DO
		fbMFunctionSpare[i].MFunction := USINT_TO_UDINT(52 + i);
		fbMFunctionSpare[i].AxesGroup := ADR(gCncXYZ);
		fbMFunctionSpare[i].Enable := TRUE;
	END_FOR

	(* Optional stop (M01) : enabled from the HMI (gCncRun.Input.OptionalStop) in Cyclic *)
	fbOptStop.AxesGroup := ADR(gCncXYZ);
	(* Start at line : velocity factor of the automatic single-axis repositioning to the start point - slow on purpose, check on site *)
	gCncRun.Input.ReposVelocityFactor := 0.1;

	(* Z reference measurement (act_MeasureZ) : own single-axis FBs. gZRef.Input (RETAIN) is kept *)
	fbZrMove[0].Axis := ADR(gAxis_X);
	fbZrMove[1].Axis := ADR(gAxis_Y);
	fbZrMove[2].Axis := ADR(gAxis_Z);
	fbZrHalt[0].Axis := ADR(gAxis_X);
	fbZrHalt[1].Axis := ADR(gAxis_Y);
	fbZrHalt[2].Axis := ADR(gAxis_Z);
	FOR i := 0 TO 2 DO
		fbZrMove[i].Acceleration := C_ZREF_ACC;
		fbZrMove[i].Deceleration := C_ZREF_ACC;
		fbZrHalt[i].Deceleration := C_ZREF_ACC;
	END_FOR
	gZRef.Output.Busy := FALSE;
	gZRef.Output.Step := 0;

	(* Work offsets G54..G57 : the active one is set as standard frame SCS1 before a run (act_WorkOffset).
	   The table (gWorkOffset, RETAIN) is kept; the axes group starts with frame 0, so woSet starts at 0 *)
	fbWorkFrame.AxesGroup := ADR(gCncXYZ);
	fbWorkFrame.CoordSystem := mcSCS1;
	fbWorkFrame.ExecutionMode := mcEM_IMMEDIATELY;
	gWorkOffset.Input.Command.Apply := FALSE;
	gWorkOffset.Output.Rejected := FALSE;
	gWorkOffset.Output.Error := FALSE;
	gWorkOffset.Output.ErrorID := 0;

	(* Head (tool) offsets : minus the mounted head's offset is set as standard frame SCS2 before a run (act_HeadOffset).
	   The table (gHeadOffset, RETAIN) is kept; the axes group starts with frame 0, so hoSet starts at 0 *)
	fbHeadFrame.AxesGroup := ADR(gCncXYZ);
	fbHeadFrame.CoordSystem := mcSCS2;
	fbHeadFrame.ExecutionMode := mcEM_IMMEDIATELY;
	gHeadOffset.Input.Command.Apply := FALSE;
	gHeadOffset.Output.Rejected := FALSE;
	gHeadOffset.Output.Error := FALSE;
	gHeadOffset.Output.ErrorID := 0;

	(* Axis reset FBs *)
	fbAxisReset[0].Axis := ADR(gAxis_X);
	fbAxisReset[1].Axis := ADR(gAxis_Y);
	fbAxisReset[2].Axis := ADR(gAxis_Z);

	(* X axis mechanical deviation compensation
	   NOTE: comp table (Position/Deviation pairs) is now defined in the axis feature
	   configuration (mcCFG_AX_FEAT_MECH_DEV_COMP) instead of runtime arrays.
	   Legacy values [mm]: P = 0 / 1000 / 2000 / 3100, D = 0 / Deviation_X1 / X2 / X3 *)
	fbMechDevCompX.Axis := ADR(gAxis_X);

	(* Teach positions C_TP1_1 .. C_TP4_3 : only CNC programs (Config_4 aliases TP1_1 ..) and the HMI (OPC UA) use them.
	   A global PV that no task references is not created on the target (OPC UA read = BadResourceUnavailable),
	   so they are referenced here once *)
	teachSum := C_TP1_1 + C_TP1_2 + C_TP1_3 + C_TP2_1 + C_TP2_2 + C_TP2_3
	          + C_TP3_1 + C_TP3_2 + C_TP3_3 + C_TP4_1 + C_TP4_2 + C_TP4_3;

END_PROGRAM
```

#### Cyclic.st - Cyclic code
```iecst
PROGRAM _CYCLIC

	(* Feedrate override from HMI *)
	IF gEquipment.Input.Parameter.Feedrate > 0.0 THEN
		fbCnc.FeedrateOverride := gEquipment.Input.Parameter.Feedrate;
	END_IF

	(* ---------- emergency stop ----------
	   MPG E-stop button, NC contact (FALSE = pressed). Software reaction only - NOT a safety circuit.
	   Stops the CNC and all single-axis motion, then powers off; discharge / laser off.
	   Latched until the button is released and RESET is sent. *)
	IF NOT DI_MPG_Jog_EMS1 THEN
		IF NOT emergencyLatched THEN
			cncCommand := E_ACT_STOP;
			commandStep := 0;
		END_IF
		emergencyLatched := TRUE;
		bootPowerDone := TRUE; (* no automatic power-on after the E-stop *)
	END_IF

	(* power on once after boot (servo only - homing is always an operator command) *)
	IF NOT bootPowerDone AND cncCommand = E_ACT_IDLE AND fbCnc.Active AND fbCnc.Info.ReadyToPowerOn THEN
		bootPowerDone := TRUE;
		initThenHome := FALSE;
		cncCommand := E_ACT_INIT;
		commandStep := 0;
	END_IF

	(* single step / optional stop (M01) from the HMI (gCncRun, both FALSE unless the HMI sets them).
	   Single step not for an MDI block (act_MoveBlock waits for MoveDone) *)
	fbCnc.SingleStep := gCncRun.Input.SingleStep AND cncCommand <> E_ACT_MOVE_BLOCK;
	fbOptStop.Enable := gCncRun.Input.OptionalStop;

	(* start at line : before its real run the program is simulated up to the start line, the axes are repositioned and it may wait for CONTINUE.
	   These phases count only in a run started by E_ACT_START_AT_LINE (lineStartRun), so START and MDI are not touched.
	   STOP, RESET, E-stop and an error end it, so an aborted start at line never blocks the next command *)
	IF cncCommand = E_ACT_STOP OR cncCommand = E_ACT_RESET OR emergencyLatched OR fbCnc.Error THEN
		lineStartRun := FALSE;
	END_IF
	lineStartPrep := lineStartRun AND fbCnc.Info.Program.ProgramPhase <> mcPRGPH_INACTIVE AND fbCnc.Info.Program.ProgramPhase <> mcPRGPH_REAL_RUN;
	lineStartWait := lineStartRun AND (fbCnc.Info.Program.ProgramPhase = mcPRGPH_WAIT_FOR_AXES_REPOS OR fbCnc.Info.Program.ProgramPhase = mcPRGPH_WAIT_FOR_REAL_RUN);

	(* program held : waits for CONTINUE - interrupted (HALT, single step), standing at M01 (fbOptStop.Interrupting is FALSE while OptionalStop is off)
	   or a start at line waiting before its real run *)
	programHeld := fbCnc.MoveInterrupted OR fbOptStop.Interrupting OR lineStartWait;

	(* program alive : running or paused (HALT). MoveActive alone is not enough - it falls on HALT,
	   so the HMI would see the run as ended and the next START would run the program from the top. A paused program counts as running everywhere below *)
	programAlive := fbCnc.MoveActive OR programHeld OR lineStartPrep;
	IF NOT programAlive AND cncCommand <> E_ACT_START_AT_LINE THEN
		lineStartRun := FALSE;
	END_IF

	(* the program stopped by itself (single step after a block, M01, start at line waiting) : act_Start leaves like after HALT so the mailbox takes CONTINUE *)
	stepHold := (fbCnc.MoveInterrupted AND fbCnc.SingleStep) OR fbOptStop.Interrupting OR lineStartWait;

	(* ---------- command preconditions ---------- *)
	CASE gEquipment.Input.CncCommand OF
		E_ACT_START: (* homing is mandatory after every power-up *)
			cmdAllowed := fbCnc.PowerOn AND fbCnc.IsHomed AND DI_Auto AND NOT programAlive;
		E_ACT_START_AT_LINE: (* like START, line 1 or later *)
			cmdAllowed := fbCnc.PowerOn AND fbCnc.IsHomed AND DI_Auto AND NOT programAlive AND gCncRun.Input.StartLine >= 1;
		E_ACT_HOME:
			cmdAllowed := fbCnc.PowerOn AND NOT programAlive;
		E_ACT_HALT:
			cmdAllowed := fbCnc.MoveActive AND NOT fbCnc.MoveInterrupted;
		E_ACT_CONTINUE: (* after HALT, a single step or M01 *)
			cmdAllowed := programHeld;
		E_ACT_POWER_OFF:
			cmdAllowed := NOT fbCnc.InMotion AND NOT programAlive;
		E_ACT_MOVE_BLOCK:
			cmdAllowed := fbCnc.PowerOn AND fbCnc.IsHomed AND NOT programAlive;
		E_ACT_MEASURE_Z: (* Z reference : manual mode, homed, every axis idle without error, no handwheel, valid gZRef.Input, sensor off *)
			cmdAllowed := fbCnc.PowerOn AND fbCnc.IsHomed AND NOT DI_Auto AND NOT programAlive AND NOT fbCnc.InMotion
				AND NOT DI_MPG_Jog_Enable AND gZRef.Output.ParamOk AND NOT DI_ZRef_Sensor
				AND gAxis[AX_X].Output.State.Status = 1 AND gAxis[AX_Y].Output.State.Status = 1 AND gAxis[AX_Z].Output.State.Status = 1;
		E_ACT_INIT, E_ACT_STOP, E_ACT_RESET, E_ACT_LOADPROGRAM:
			cmdAllowed := TRUE;
		ELSE (* a value without an action (ABORT while idle, unknown) : refused, so it never blocks the mailbox *)
			cmdAllowed := FALSE;
	END_CASE

	(* during an E-stop only STOP / RESET / servo off are accepted *)
	IF emergencyLatched AND gEquipment.Input.CncCommand <> E_ACT_STOP AND gEquipment.Input.CncCommand <> E_ACT_RESET AND gEquipment.Input.CncCommand <> E_ACT_POWER_OFF THEN
		cmdAllowed := FALSE;
	END_IF

	(* ---------- command arbitration ---------- *)
	IF cncCommand <> gEquipment.Input.CncCommand AND cncCommand = E_ACT_IDLE THEN

		IF cmdAllowed THEN

			cncCommand := gEquipment.Input.CncCommand;
			initThenHome := TRUE; (* INIT from HMI = power + homing *)
			gEquipment.Output.Status.Rejected := E_ACT_IDLE;
			gEquipment.Input.CncCommand := E_ACT_IDLE;
			commandStep := 0;
		ELSE
			gEquipment.Output.Status.Rejected := gEquipment.Input.CncCommand;
			gEquipment.Input.CncCommand := E_ACT_IDLE;
		END_IF

	ELSIF gEquipment.Input.CncCommand = E_ACT_HALT AND cmdAllowed AND (cncCommand = E_ACT_START OR cncCommand = E_ACT_CONTINUE OR cncCommand = E_ACT_START_AT_LINE) THEN

		cncCommand := gEquipment.Input.CncCommand;
		gEquipment.Input.CncCommand := E_ACT_IDLE;
		commandStep := 0;

	ELSIF gEquipment.Input.CncCommand = E_ACT_STOP AND cncCommand <> E_ACT_IDLE AND cncCommand <> E_ACT_INIT THEN

		cncCommand := gEquipment.Input.CncCommand;
		gEquipment.Input.CncCommand := E_ACT_IDLE;
		commandStep := 0;

	ELSIF cncCommand <> E_ACT_IDLE AND gEquipment.Input.CncCommand = E_ACT_ABORT THEN

		gEquipment.Input.CncCommand := E_ACT_IDLE;
		cncCommand := E_ACT_IDLE;

	ELSIF cncCommand <> E_ACT_IDLE THEN

		gEquipment.Input.CncCommand := E_ACT_IDLE;

	END_IF

	(* work offset G54..G57 : Apply from the HMI, frame SCS1 set before a run (only when an offset is in use) *)
	act_WorkOffset;

	(* head offset : Apply from the HMI, frame SCS2 set before a run (only when an offset is in use) *)
	act_HeadOffset;

	(* program start point : from the top (the B&R defaults), except while E_ACT_START_AT_LINE starts a program (act_Start step 0),
	   so START and MDI never inherit a start line through fbCnc.Update *)
	IF cncCommand <> E_ACT_START_AT_LINE THEN
		CncParameters.MoveProgramOptions.StartPointType := mcPRGSP_STANDARD;
		CncParameters.MoveProgramOptions.StartPointParameter := 0.0;
		CncParameters.MoveProgramOptions.RepositioningParameter.Type := mcPRGRP_SINGLE_AXIS;
		CncParameters.MoveProgramOptions.RepositioningParameter.AxisVelocityFactor := 0.0;
	END_IF

	(* ---------- command execution ---------- *)
	CASE cncCommand OF

		E_ACT_IDLE:

			commandStep := 0;

			(* release all pulse-type CNC commands - MoveProgram only once the program has ended : a paused program must stay loaded for CONTINUE *)
			fbCnc.Home := FALSE;
			IF NOT programAlive THEN
				fbCnc.MoveProgram := FALSE;
			END_IF
			fbCnc.MoveBlock := FALSE;
			fbCnc.Interrupt := FALSE;
			fbCnc.Continue := FALSE;
			fbOptStop.Continue := FALSE;
			fbCnc.Stop := FALSE;
			fbCnc.ErrorReset := FALSE;
			fbCnc.Update := FALSE;
			fbAxisReset[0].Execute := FALSE;
			fbAxisReset[1].Execute := FALSE;
			fbAxisReset[2].Execute := FALSE;

			stepTimer(IN := FALSE);

		E_ACT_INIT:

			act_Init;

			IF commandStep = 100 THEN
				commandStep := 0;
				IF initThenHome AND NOT fbCnc.IsHomed THEN
					cncCommand := E_ACT_HOME;
				ELSE
					cncCommand := E_ACT_IDLE;
				END_IF
			ELSIF commandStep = 200 THEN
				cncCommand := E_ACT_IDLE;
			END_IF

		E_ACT_LOADPROGRAM: (* Load CNC Program *)

			cncCommand := E_ACT_IDLE;

		E_ACT_START: (* Execute CNC *)

			act_Start;

			IF commandStep = 100 THEN
				cncCommand := E_ACT_IDLE;
			ELSIF commandStep = 200 THEN
				cncCommand := E_ACT_IDLE;
			END_IF

		E_ACT_START_AT_LINE: (* Execute CNC from the file line gCncRun.Input.StartLine - act_Start sets the start point *)

			act_Start;

			IF commandStep = 100 OR commandStep = 200 THEN
				cncCommand := E_ACT_IDLE;
			END_IF

		E_ACT_RESET: (* CNC Reset *)

			act_Reset;

			IF commandStep = 100 OR commandStep = 200 THEN
				cncCommand := E_ACT_IDLE;
			END_IF

		E_ACT_HOME:

			IF NOT fbCnc.InMotion THEN
				act_Home;
			END_IF

			IF commandStep = 100 OR commandStep = 200 THEN
				cncCommand := E_ACT_IDLE;
			END_IF

		E_ACT_HALT: (* CNC Halt *)

			act_Halt;

			IF commandStep = 2 THEN
				commandStep := 0;
				cncCommand := E_ACT_IDLE;
			END_IF

		E_ACT_CONTINUE: (* CNC Continue *)

			act_Continue;

			IF commandStep = 1 THEN
				commandStep := 0;
				cncCommand := E_ACT_IDLE;
			END_IF

		E_ACT_STOP: (* CNC Stop *)

			act_Stop;

			IF commandStep = 2 THEN
				commandStep := 0;
				cncCommand := E_ACT_IDLE;
			END_IF

		E_ACT_POWER_OFF: (* Servo off *)

			act_PowerOff;

			IF commandStep = 100 OR commandStep = 200 THEN
				cncCommand := E_ACT_IDLE;
			END_IF

		E_ACT_MOVE_BLOCK: (* MDI : single NC block *)

			act_MoveBlock;

			IF commandStep = 100 OR commandStep = 200 THEN
				cncCommand := E_ACT_IDLE;
			END_IF

		E_ACT_MEASURE_Z: (* Z reference measurement : result in gZRef.Output *)

			act_MeasureZ;

			IF commandStep = 100 OR commandStep = 200 THEN
				cncCommand := E_ACT_IDLE;
			END_IF

	END_CASE

	(* Z reference : input check, a measurement left by STOP / ABORT / E-stop / handwheel is braked, status *)
	act_ZRef;

	(* program finished : also after HALT / CONTINUE, when act_Start is no longer running and cannot see MoveDone.
	   The program ends without STOP, error or interruption -> Complete *)
	programEndTrig(CLK := programAlive);
	IF programEndTrig.Q AND programStarted THEN
		IF NOT fbCnc.Error AND NOT fbCnc.MoveInterrupted AND NOT gEquipment.Output.State.Stop THEN
			gEquipment.Output.State.Complete := TRUE;
		END_IF
		programStarted := FALSE;
	END_IF

	(* LaserPower set by a program or an MDI line (path synchronous alias) holds for that run only *)
	IF programEndTrig.Q THEN
		C_LaserPower := -1.0;
	END_IF

	(* E-stop : power off once the axes have stopped (at the latest after 2 s) *)
	emergencyTimer(IN := emergencyLatched, PT := T#2s);
	IF emergencyLatched AND (NOT fbCnc.InMotion OR emergencyTimer.Q) THEN
		fbCnc.Power := FALSE;
	END_IF

	(* ---------- status to HMI ---------- *)
	gEquipment.Output.Status.CurrentAction := cncCommand;
	gEquipment.Output.Status.Mode := DI_Auto;
	gEquipment.Output.State.Move := fbCnc.InMotion;
	gEquipment.Output.Status.PowerOn := fbCnc.PowerOn;
	gEquipment.Output.Status.IsHomed := fbCnc.IsHomed;
	gEquipment.Output.Status.ProgramActive := programAlive; (* TRUE while paused too - HMI, OpMode, AxisManual (idle), Laser read it *)
	gEquipment.Output.Status.ProgramInterrupted := programHeld; (* HALT, single step or M01 : the HMI offers CONTINUE *)
	gEquipment.Output.Status.Error := fbCnc.Error;
	gEquipment.Output.Status.StatusID := fbCnc.StatusID;
	gEquipment.Output.Status.EmergencyStop := emergencyLatched;
	C_CurrentLine := UDINT_TO_DINT(fbCnc.Info.Program.ProgramMonitor.LineNumber);
	C_OverallRuntime := fbCnc.Info.Program.ProgramMonitor.OverallRuntime; (* HMI : remaining time, elapsed time *)
	C_MovementRuntime := fbCnc.Info.Program.ProgramMonitor.MovementRuntime;
	gHeadSupport := SHL(UDINT#1, HEAD_DISPENSER) OR SHL(UDINT#1, HEAD_LASER); (* heads of this PLC program - fixed, set every cycle so a write over OPC UA does not stay *)
	gCncRun.Output.SingleStepActive := fbCnc.SingleStepActive;
	gCncRun.Output.OptionalStopActive := fbOptStop.Interrupting;
	gCncRun.Output.OptionalStopErrorId := fbOptStop.ErrorID;
	gCncRun.Output.InterruptStatus := fbCnc.Info.Program.InterruptStatus;
	gCncRun.Output.ProgramPhase := fbCnc.Info.Program.ProgramPhase;

	(* ---------- M functions ---------- *)
	mfClear := NOT programAlive OR emergencyLatched; (* no program / E-stop : M42, M62 act as if set - not while paused, M41 / M61 come back after CONTINUE *)

	act_HeadCheck; (* only the M functions and manual on of the active head (gActiveHead) - 0 = no check *)

	act_M41;
	act_M42;
	act_M44;
	act_M45;
	act_MSpare; (* M50..M59 : no function, go on at once *)
	act_M61;
	act_M62;

	(* HALT, single step, M01 : output off while the program is held, back on after CONTINUE (M41 / M61 Value stays set) *)
	IF programHeld THEN
		gDispenser.Input.Command.Discharge := FALSE;
		gLaser.Input.Command.Emission := FALSE;
	END_IF

	IF emergencyLatched THEN
		gDispenser.Input.Command.Manual := FALSE;
		gLaser.Input.Command.Manual := FALSE;
	END_IF

	(* ---------- FB calls ---------- *)
	fbCnc();
	fbOptStop();

	FOR i := 0 TO 7 DO
		fbMFunction[i]();
		fbMFunctionSpare[i]();
	END_FOR

	FOR i := 0 TO 2 DO
		fbAxisReset[i]();
	END_FOR

	fbMechDevCompX();

	FOR i := 0 TO 2 DO
		fbZrMove[i]();
		fbZrHalt[i]();
	END_FOR
	fbWorkFrame();
	fbHeadFrame();

END_PROGRAM
```

#### Exit.st - Exit code
```iecst
PROGRAM _EXIT
END_PROGRAM
```

#### Action_NC.st - NC actions
```iecst
ACTION act_Halt:

	CASE commandStep OF
		0:
			fbCnc.Interrupt := TRUE;
			commandStep := 1;
		1:
			IF fbCnc.MoveInterrupted = TRUE THEN
				fbCnc.Interrupt := FALSE;
				commandStep := 2;
			END_IF
		2:
			;(* Complete *)
	END_CASE
END_ACTION

ACTION act_Stop:

	CASE commandStep OF
		0:
			gEquipment.Output.State.Stop := TRUE;
			programStarted := FALSE;
			fbCnc.Stop := fbCnc.PowerOn; (* nothing to stop without power *)
			commandStep := 1;
		1:
			IF fbCnc.InMotion = FALSE THEN
				fbCnc.Stop := FALSE;
				commandStep := 2;
			END_IF
		2:
			;(* Complete *)
	END_CASE
END_ACTION

ACTION act_Init:
	CASE commandStep OF
		0:
			stepTimer(IN := FALSE);

			IF fbCnc.Active = TRUE AND fbCnc.Info.CommunicationReady = TRUE THEN
				commandStep := 5;
			END_IF

		5:
			(* Power is level-sensitive and needs a new rising edge after an error : drop it for one cycle *)
			IF fbCnc.PowerOn = TRUE THEN
				commandStep := 100;
			ELSE
				fbCnc.Power := FALSE;
				commandStep := 10;
			END_IF

		10:
			fbCnc.Power := TRUE; (* powers all group axes *)
			stepTimer(IN := TRUE, PT := T#10s);

			IF fbCnc.PowerOn = TRUE THEN
				stepTimer(IN := FALSE);
				commandStep := 100;
			ELSIF fbCnc.Error OR stepTimer.Q THEN
				stepTimer(IN := FALSE);
				fbCnc.Power := FALSE;
				commandStep := 200;
			END_IF

		100:
			;(* Complete *)

		200:
			;(* power on failed - see gEquipment.Output.Status.Error / StatusID *)
	END_CASE
END_ACTION

ACTION act_Reset:
	CASE commandStep OF
		0:
			(* E-stop is cleared only once the button is released *)
			IF DI_MPG_Jog_EMS1 THEN
				emergencyLatched := FALSE;
			END_IF

			fbCnc.ErrorReset := TRUE;

			fbAxisReset[0].Execute := TRUE;
			fbAxisReset[1].Execute := TRUE;
			fbAxisReset[2].Execute := TRUE;

			commandStep := 10;

		10:
			IF NOT fbAxisReset[0].Busy AND NOT fbAxisReset[1].Busy AND NOT fbAxisReset[2].Busy THEN
				commandStep := 20;
			END_IF

		20:
			fbCnc.ErrorReset := FALSE;
			fbAxisReset[0].Execute := FALSE;
			fbAxisReset[1].Execute := FALSE;
			fbAxisReset[2].Execute := FALSE;
			stepTimer(IN := TRUE, PT := T#3s);

			IF fbCnc.Error = FALSE THEN
				stepTimer(IN := FALSE);
				commandStep := 100;
			ELSIF stepTimer.Q THEN
				(* error cause still present *)
				stepTimer(IN := FALSE);
				commandStep := 200;
			END_IF
		100:
			;(* Complete - servo stays off after an error : operator sends INIT *)
		200:
			;(* reset failed *)
	END_CASE
END_ACTION

ACTION act_Continue:
	CASE commandStep OF
		0:
			IF fbOptStop.Interrupting THEN
				fbOptStop.Continue := TRUE; (* standing at M01 - released in IDLE like fbCnc.Continue *)
			ELSIF fbCnc.MoveInterrupted OR lineStartWait THEN
				fbCnc.Continue := TRUE; (* HALT, single step : next block. Start at line : reposition / real run *)
			END_IF
			commandStep := 1;
		1:
			IF NOT fbCnc.MoveInterrupted THEN
				fbCnc.Continue := FALSE;
			END_IF
	END_CASE
END_ACTION

ACTION act_Home:
	CASE commandStep OF
		0:
			(* homing mode / home offsets are defined in the axis homing configuration. *)
			gEquipment.Output.State.Initialized := FALSE;

			IF fbCnc.PowerOn THEN
				fbCnc.Home := TRUE;
				commandStep := 5;
			ELSE
				commandStep := 200;
			END_IF

		5:
			IF fbCnc.CommandBusy = TRUE THEN
				commandStep := 10;
			ELSIF fbCnc.Error OR fbCnc.CommandAborted THEN
				fbCnc.Home := FALSE;
				commandStep := 200;
			END_IF

		10:
			IF fbCnc.IsHomed = TRUE AND fbCnc.CommandBusy = FALSE THEN
				fbCnc.Home := FALSE;
				commandStep := 20;
			ELSIF fbCnc.Error OR fbCnc.CommandAborted OR (fbCnc.CommandBusy = FALSE AND fbCnc.IsHomed = FALSE) THEN
				fbCnc.Home := FALSE;
				commandStep := 200;
			END_IF

		20:
			(* X axis mechanical deviation compensation - table from axis feature config *)
			fbMechDevCompX.Command := mcMDC_CMD_SWITCH_ON;
			fbMechDevCompX.Execute := TRUE;

			IF fbMechDevCompX.Done THEN
				fbMechDevCompX.Execute := FALSE;
				commandStep := 30;
			ELSIF fbMechDevCompX.Error THEN
				(* compensation feature not configured -> continue without it *)
				fbMechDevCompX.Execute := FALSE;
				commandStep := 30;
			END_IF

		30:
			(* a wait position after homing is up to the HMI (ManualPositon + ManualMove) *)
			commandStep := 50;

		50:
			gEquipment.Input.Command.AlarmClearAll := TRUE;
			gEquipment.Output.State.Initialized := TRUE;
			commandStep := 100;

		100:
			;

		200:
			;(* homing failed or servo off *)
	END_CASE
END_ACTION

ACTION act_Start:

	CASE commandStep OF
		0:
			stepTimer(IN := FALSE);
			gEquipment.Output.Status.WorkPanelName := gEquipment.Input.Parameter.sProgramName;
			CncParameters.ProgramName := gEquipment.Input.Parameter.sProgramName;
			CncParameters.MoveProgramOptions.InitProgram := gEquipment.Input.Parameter.sInitProgram;
			IF cncCommand = E_ACT_START_AT_LINE THEN
				(* start at the file line StartLine (1 = first, as C_CurrentLine) : mapp simulates the program up to that line, then moves
				   the axes to its start point by itself with single-axis moves. Cyclic puts the standard start point back once 15 is over *)
				CncParameters.MoveProgramOptions.StartPointType := mcPRGSP_LINE_NUMBER;
				CncParameters.MoveProgramOptions.StartPointParameter := UDINT_TO_LREAL(gCncRun.Input.StartLine);
				CncParameters.MoveProgramOptions.RepositioningParameter.Type := mcPRGRP_SINGLE_AXIS_AUTOMATIC;
				CncParameters.MoveProgramOptions.RepositioningParameter.AxisVelocityFactor := gCncRun.Input.ReposVelocityFactor;
			END_IF
			fbCnc.Update := TRUE;
			commandStep := 1;

		1:
			stepTimer(IN := TRUE, PT := T#5s);

			IF fbCnc.UpdateDone = TRUE THEN
				fbCnc.Update := FALSE;
				commandStep := 2;
			ELSIF stepTimer.Q THEN
				stepTimer(IN := FALSE);
				fbCnc.Update := FALSE;
				commandStep := 200;
			END_IF

		2:
			gEquipment.Output.State.Stop := FALSE;
			gEquipment.Output.State.Complete := FALSE;
			IF woNeed THEN
				(* work offset in use : set its frame first (act_WorkOffset) *)
				woStep := 1;
				commandStep := 5;
			ELSIF hoNeed THEN
				(* head offset in use : set its frame first (act_HeadOffset) *)
				hoStep := 1;
				commandStep := 6;
			ELSE
				commandStep := 10;
			END_IF

		5:
			IF woStep = 100 THEN
				IF hoNeed THEN
					(* head offset in use too : set its frame next (act_HeadOffset) *)
					hoStep := 1;
					commandStep := 6;
				ELSE
					commandStep := 10;
				END_IF
			ELSIF woStep = 200 THEN
				commandStep := 200; (* gWorkOffset.Output.Error / ErrorID *)
			END_IF

		6:
			IF hoStep = 100 THEN
				commandStep := 10;
			ELSIF hoStep = 200 THEN
				commandStep := 200; (* gHeadOffset.Output.Error / ErrorID *)
			END_IF

		10:
			fbCnc.MoveProgram := TRUE;
			programStarted := TRUE;
			lineStartRun := cncCommand = E_ACT_START_AT_LINE; (* FALSE for START *)
			commandStep := 20;

		20:
			IF fbCnc.MoveActive = TRUE THEN
				commandStep := 30;
			ELSIF fbCnc.Error = TRUE THEN
				fbCnc.MoveProgram := FALSE;
				commandStep := 200;
			ELSIF stepHold THEN
				(* single step / M01 / start at line waiting stopped the program before MoveActive was seen - see step 30 *)
				commandStep := 100;
			END_IF

		30:
			IF fbCnc.MoveDone = TRUE THEN
				fbCnc.MoveProgram := FALSE;
				gEquipment.Output.State.Complete := TRUE;
				commandStep := 100;
			ELSIF fbCnc.Error OR fbCnc.CommandAborted THEN
				(* program error / aborted while running *)
				fbCnc.MoveProgram := FALSE;
				commandStep := 200;
			ELSIF stepHold THEN
				(* single step / M01 / start at line waiting : the program waits for CONTINUE. Leave like after HALT so the mailbox takes CONTINUE -
				   MoveProgram stays set while the program is alive (IDLE branch), programEndTrig reports Complete at the end *)
				commandStep := 100;
			END_IF

		100:
			;(* Complete *)

		200:
			;(* load / start error *)
	END_CASE

END_ACTION

ACTION act_PowerOff:

	CASE commandStep OF
		0:
			stepTimer(IN := FALSE);
			fbCnc.Power := FALSE;
			commandStep := 10;

		10:
			stepTimer(IN := TRUE, PT := T#5s);

			IF fbCnc.PowerOn = FALSE THEN
				stepTimer(IN := FALSE);
				commandStep := 100;
			ELSIF stepTimer.Q THEN
				stepTimer(IN := FALSE);
				commandStep := 200;
			END_IF

		100:
			;(* Complete *)

		200:
			;(* servo did not switch off *)
	END_CASE

END_ACTION

ACTION act_MoveBlock:

	CASE commandStep OF
		0:
			stepTimer(IN := FALSE);
			programStarted := FALSE; (* an MDI block is not a production run *)
			CncParameters.Block := gEquipment.Input.Parameter.sBlock;
			fbCnc.Update := TRUE;
			commandStep := 1;

		1:
			stepTimer(IN := TRUE, PT := T#5s);

			IF fbCnc.UpdateDone = TRUE THEN
				stepTimer(IN := FALSE);
				fbCnc.Update := FALSE;
				IF woNeed THEN
					(* work offset in use : set its frame first (act_WorkOffset) *)
					woStep := 1;
					commandStep := 5;
				ELSIF hoNeed THEN
					(* head offset in use : set its frame first (act_HeadOffset) *)
					hoStep := 1;
					commandStep := 6;
				ELSE
					commandStep := 10;
				END_IF
			ELSIF stepTimer.Q THEN
				stepTimer(IN := FALSE);
				fbCnc.Update := FALSE;
				commandStep := 200;
			END_IF

		5:
			IF woStep = 100 THEN
				IF hoNeed THEN
					(* head offset in use too : set its frame next (act_HeadOffset) *)
					hoStep := 1;
					commandStep := 6;
				ELSE
					commandStep := 10;
				END_IF
			ELSIF woStep = 200 THEN
				commandStep := 200; (* gWorkOffset.Output.Error / ErrorID *)
			END_IF

		6:
			IF hoStep = 100 THEN
				commandStep := 10;
			ELSIF hoStep = 200 THEN
				commandStep := 200; (* gHeadOffset.Output.Error / ErrorID *)
			END_IF

		10:
			gEquipment.Output.State.Complete := FALSE;
			(* MoveDone / CommandAborted still set by an earlier move (e.g. a program that ended after HALT / CONTINUE,
			   when MoveProgram was already FALSE) are not this block's - step 20 ignores them until they fall *)
			mdiDoneOld := fbCnc.MoveDone;
			mdiAbortOld := fbCnc.CommandAborted;
			fbCnc.MoveBlock := TRUE;
			commandStep := 20;

		20:
			(* like act_Start : running first, then done. Not started within 5 s -> failed *)
			stepTimer(IN := TRUE, PT := T#5s);

			IF NOT fbCnc.MoveDone THEN
				mdiDoneOld := FALSE;
			END_IF
			IF NOT fbCnc.CommandAborted THEN
				mdiAbortOld := FALSE;
			END_IF

			IF fbCnc.MoveActive = TRUE THEN
				stepTimer(IN := FALSE);
				commandStep := 30;
			ELSIF fbCnc.MoveDone = TRUE AND NOT mdiDoneOld THEN
				(* short block already finished *)
				stepTimer(IN := FALSE);
				fbCnc.MoveBlock := FALSE;
				commandStep := 100;
			ELSIF fbCnc.Error OR (fbCnc.CommandAborted AND NOT mdiAbortOld) THEN
				stepTimer(IN := FALSE);
				fbCnc.MoveBlock := FALSE;
				commandStep := 200;
			ELSIF stepTimer.Q THEN
				stepTimer(IN := FALSE);
				fbCnc.MoveBlock := FALSE;
				commandStep := 200;
			END_IF

		30:
			IF fbCnc.MoveDone = TRUE THEN
				fbCnc.MoveBlock := FALSE;
				commandStep := 100;
			ELSIF fbCnc.Error OR fbCnc.CommandAborted THEN
				fbCnc.MoveBlock := FALSE;
				commandStep := 200;
			END_IF

		100:
			;(* Complete *)

		200:
			;(* block rejected or failed - see Output.Status.Error / StatusID *)
	END_CASE

END_ACTION
```

#### Action_MCode.st - M-code actions
```iecst
(* Nozzle Valve Open *)
ACTION act_M41: (* Asynchronous *)

	IF fbMFunction[0].Value = TRUE AND headDispOk THEN (* another head active : refused in act_HeadCheck *)
		gDispenser.Input.Command.Discharge := TRUE;
		fbMFunction[1].Reset := TRUE; (* on/off pair : M41 clears the latched M42 and M42 clears M41, so the last one holds *)
	ELSE
		fbMFunction[1].Reset := FALSE;
	END_IF

END_ACTION

(* Nozzle Valve Close - also while no program runs / E-stop (mfClear), so M41 does not stay on *)
ACTION act_M42: (* Asynchronous *)

	IF fbMFunction[1].Value = TRUE OR mfClear THEN
		gDispenser.Input.Command.Discharge := FALSE;
		fbMFunction[0].Reset := TRUE;
	ELSE
		fbMFunction[0].Reset := FALSE;
	END_IF

END_ACTION

(* Valve Delay On *)
ACTION act_M44: (* Asynchronous *)

	IF fbMFunction[2].Value = TRUE THEN
		gDispenser.Input.Parameter.DischargeDelay := TRUE;
		fbMFunction[2].Reset := TRUE;
	ELSE
		fbMFunction[2].Reset := FALSE;
	END_IF

END_ACTION

(* Valve Delay Off *)
ACTION act_M45: (* Asynchronous *)

	IF fbMFunction[3].Value = TRUE THEN
		gDispenser.Input.Parameter.DischargeDelay := FALSE;
		fbMFunction[3].Reset := TRUE;
	ELSE
		fbMFunction[3].Reset := FALSE;
	END_IF

END_ACTION

(* M50..M59 (blocking, range 50..59 of the axes group M-function feature) : no function on this machine. Without a handler the path
   would wait at such a line for ever - reset at once, the program goes on as if the line were not there.
   fbMFunction[6] / [7] watch M50 / M51, fbMFunctionSpare[0..7] M52..M59 *)
ACTION act_MSpare: (* Synchronous *)

	FOR i := 6 TO 7 DO
		IF fbMFunction[i].Value = TRUE THEN
			fbMFunction[i].Reset := TRUE;
			mfSpareLast := 44 + i;
		ELSE
			fbMFunction[i].Reset := FALSE;
		END_IF
	END_FOR

	FOR i := 0 TO 7 DO
		IF fbMFunctionSpare[i].Value = TRUE THEN
			fbMFunctionSpare[i].Reset := TRUE;
			mfSpareLast := 52 + i;
		ELSE
			fbMFunctionSpare[i].Reset := FALSE;
		END_IF
	END_FOR

END_ACTION

(* Laser On *)
ACTION act_M61: (* Asynchronous *)

	IF fbMFunction[4].Value = TRUE AND headLaserOk THEN (* another head active : refused in act_HeadCheck *)
		gLaser.Input.Command.Emission := TRUE;
		fbMFunction[5].Reset := TRUE; (* on/off pair, as M41 / M42 *)
	ELSE
		fbMFunction[5].Reset := FALSE;
	END_IF

END_ACTION

(* Laser Off - also while no program runs / E-stop (mfClear), so M61 does not stay on *)
ACTION act_M62: (* Asynchronous *)

	IF fbMFunction[5].Value = TRUE OR mfClear THEN
		gLaser.Input.Command.Emission := FALSE;
		fbMFunction[4].Reset := TRUE;
	ELSE
		fbMFunction[4].Reset := FALSE;
	END_IF

END_ACTION
```

#### Action_Head.st - Head actions
```iecst
(* One head on the machine (HMI plugin structure). Head number HEAD_* = PlcId of the HMI head plugin.
   gActiveHead (written by the HMI) : only the M functions and the manual on of that head are taken. An M function of another head
   stops the running program (like STOP from the HMI : the run ends as stopped, not complete), a manual on of another head is dropped,
   its outputs stay off; gHeadRefused shows that head until the next run starts or RESET.
   gActiveHead = 0 (not written yet after a PLC restart) : no check *)
ACTION act_HeadCheck:

	headDispOk := gActiveHead = 0 OR gActiveHead = HEAD_DISPENSER;
	headLaserOk := gActiveHead = 0 OR gActiveHead = HEAD_LASER;

	(* the last refusal shows until the next run starts or RESET *)
	headRunTrig(CLK := programAlive);
	IF headRunTrig.Q OR cncCommand = E_ACT_RESET THEN
		gHeadRefused := 0;
	END_IF

	(* an on code (M41 / M61) counts by its value - it is held in reset while no program runs (mfClear, act_M42 / act_M62).
	   The off codes (M42 / M62, reset only by the next on code) and the delay flags (M44 / M45, pulses) count on their rising edge,
	   so a value left over from an earlier run of the other head is not taken as new *)
	FOR i := 0 TO 5 DO
		headMfTrig[i](CLK := fbMFunction[i].Value);
	END_FOR

	headRefuse := 0;
	IF NOT headDispOk AND (fbMFunction[0].Value OR headMfTrig[1].Q OR headMfTrig[2].Q OR headMfTrig[3].Q) THEN
		headRefuse := HEAD_DISPENSER;
	END_IF
	IF NOT headLaserOk AND (fbMFunction[4].Value OR headMfTrig[5].Q) THEN
		headRefuse := HEAD_LASER;
	END_IF

	IF headRefuse <> 0 THEN
		gHeadRefused := headRefuse;
		IF programAlive AND cncCommand <> E_ACT_STOP THEN
			cncCommand := E_ACT_STOP;
			commandStep := 0;
		END_IF
	END_IF

	(* a head that is not the active one stays off : act_M41 / act_M61 do not switch it on, its manual on is dropped *)
	IF NOT headDispOk THEN
		IF gDispenser.Input.Command.Manual THEN
			gHeadRefused := HEAD_DISPENSER;
		END_IF
		gDispenser.Input.Command.Discharge := FALSE;
		gDispenser.Input.Command.Manual := FALSE;
	END_IF

	IF NOT headLaserOk THEN
		IF gLaser.Input.Command.Manual THEN
			gHeadRefused := HEAD_LASER;
		END_IF
		gLaser.Input.Command.Emission := FALSE;
		gLaser.Input.Command.Manual := FALSE;
	END_IF

END_ACTION
```

#### Action_ZRef.st - Z reference measurement actions
```iecst
ACTION act_ZRefCheck:
	(* gZRef.Input valid for a measurement (machine coordinates, Z+ down, 0 = top) : SafeZ <= StartZ < MaxZ, search at most
	   C_ZREF_MAX_SEARCH, everything inside the software limits of gAxis[].Input.Parameter (loaded from the axis configuration
	   by AxisManual), search velocity at most C_ZREF_MAX_VEL. The defaults (all 0) are not valid : nothing moves until the HMI
	   has written the sensor position *)
	zrVel := gZRef.Input.ProbeVel;
	IF zrVel <= 0.0 THEN
		zrVel := C_ZREF_PROBE_VEL;
	END_IF

	gZRef.Output.ParamOk := gZRef.Input.MaxZ > gZRef.Input.StartZ
		AND gZRef.Input.MaxZ - gZRef.Input.StartZ <= C_ZREF_MAX_SEARCH
		AND gZRef.Input.SafeZ <= gZRef.Input.StartZ
		AND zrVel <= C_ZREF_MAX_VEL
		AND gZRef.Input.SafeZ >= DINT_TO_LREAL(gAxis[AX_Z].Input.Parameter.SoftwareLimitsNeg)
		AND gZRef.Input.MaxZ <= DINT_TO_LREAL(gAxis[AX_Z].Input.Parameter.SoftwareLimitsPos)
		AND gZRef.Input.SensorX >= DINT_TO_LREAL(gAxis[AX_X].Input.Parameter.SoftwareLimitsNeg)
		AND gZRef.Input.SensorX <= DINT_TO_LREAL(gAxis[AX_X].Input.Parameter.SoftwareLimitsPos)
		AND gZRef.Input.SensorY >= DINT_TO_LREAL(gAxis[AX_Y].Input.Parameter.SoftwareLimitsNeg)
		AND gZRef.Input.SensorY <= DINT_TO_LREAL(gAxis[AX_Y].Input.Parameter.SoftwareLimitsPos);

END_ACTION

ACTION act_MeasureZ:
	(* Z reference measurement (CncCommand E_ACT_MEASURE_Z) : Z up to SafeZ, X / Y to the sensor, Z to StartZ, then Z slowly
	   down towards MaxZ until the touch sensor DI_ZRef_Sensor comes on : that Z is the result (gZRef.Output.MeasuredZ, the
	   HMI puts it into the head table), Z brakes and goes back up to SafeZ. Single-axis moves in machine coordinates with
	   own FBs (fbZrMove / fbZrHalt), like AxisManual's ManualMove; the CNC program path is not used, so work / head offsets
	   do not shift it. Accepted only in manual mode, homed, standing (preconditions in Cyclic).
	   DI_ZRef_Sensor is NOT wired yet : without a sensor the search reaches MaxZ and ends with ErrorId 3 *)

	CASE commandStep OF
		0: (* take the input over, clear the last result *)
			stepTimer(IN := FALSE);
			act_ZRefCheck;
			gZRef.Output.Done := FALSE;
			gZRef.Output.ErrorId := 0;
			zrFail := 0;
			FOR i := 0 TO 2 DO
				fbZrMove[i].Execute := FALSE;
				fbZrHalt[i].Execute := FALSE;
			END_FOR
			zrMoveVel := gEquipment.Input.Parameter.SystemSpeed; (* like ManualMove *)
			IF zrMoveVel <= 0.0 THEN
				zrMoveVel := C_ZREF_MOVE_VEL;
			END_IF

			IF gZRef.Output.ParamOk THEN
				zrActive := TRUE;
				commandStep := 10;
			ELSE
				gZRef.Output.ErrorId := 1;
				commandStep := 200;
			END_IF

		10: (* Z up to SafeZ first - a head already above SafeZ stays there (Z never goes down before X / Y move) *)
			fbZrMove[2].Position := MIN(gZRef.Input.SafeZ, gAxis[AX_Z].Output.State.Position);
			fbZrMove[2].Velocity := zrMoveVel;
			fbZrMove[2].Execute := TRUE;
			stepTimer(IN := FALSE);
			commandStep := 11;

		11:
			stepTimer(IN := TRUE, PT := T#60s);

			IF fbZrMove[2].Done THEN
				stepTimer(IN := FALSE);
				fbZrMove[2].Execute := FALSE;
				commandStep := 20;
			ELSIF fbZrMove[2].Error OR fbZrMove[2].CommandAborted THEN
				zrFail := 4;
				commandStep := 190;
			ELSIF stepTimer.Q THEN
				zrFail := 6;
				commandStep := 190;
			END_IF

		20: (* X / Y over the sensor *)
			fbZrMove[0].Position := gZRef.Input.SensorX;
			fbZrMove[0].Velocity := zrMoveVel;
			fbZrMove[0].Execute := TRUE;
			fbZrMove[1].Position := gZRef.Input.SensorY;
			fbZrMove[1].Velocity := zrMoveVel;
			fbZrMove[1].Execute := TRUE;
			stepTimer(IN := FALSE);
			commandStep := 21;

		21:
			stepTimer(IN := TRUE, PT := T#60s);

			IF fbZrMove[0].Done AND fbZrMove[1].Done THEN
				stepTimer(IN := FALSE);
				fbZrMove[0].Execute := FALSE;
				fbZrMove[1].Execute := FALSE;
				commandStep := 30;
			ELSIF fbZrMove[0].Error OR fbZrMove[0].CommandAborted OR fbZrMove[1].Error OR fbZrMove[1].CommandAborted THEN
				zrFail := 4;
				commandStep := 190;
			ELSIF stepTimer.Q THEN
				zrFail := 6;
				commandStep := 190;
			END_IF

		30: (* Z down to StartZ *)
			fbZrMove[2].Position := gZRef.Input.StartZ;
			fbZrMove[2].Velocity := zrMoveVel;
			fbZrMove[2].Execute := TRUE;
			stepTimer(IN := FALSE);
			commandStep := 31;

		31:
			stepTimer(IN := TRUE, PT := T#60s);

			IF fbZrMove[2].Done THEN
				stepTimer(IN := FALSE);
				fbZrMove[2].Execute := FALSE;
				commandStep := 40;
			ELSIF fbZrMove[2].Error OR fbZrMove[2].CommandAborted THEN
				zrFail := 4;
				commandStep := 190;
			ELSIF stepTimer.Q THEN
				zrFail := 6;
				commandStep := 190;
			END_IF

		40: (* slow search towards MaxZ - the sensor must be off here (else StartZ is too low or the sensor is stuck) *)
			IF DI_ZRef_Sensor THEN
				zrFail := 2;
				commandStep := 60;
			ELSE
				fbZrMove[2].Position := gZRef.Input.MaxZ;
				fbZrMove[2].Velocity := zrVel;
				fbZrMove[2].Execute := TRUE;
				stepTimer(IN := FALSE);
				commandStep := 41;
			END_IF

		41:
			stepTimer(IN := TRUE, PT := T#60s);

			IF DI_ZRef_Sensor THEN
				(* Z of the last cycle (AxisManual runs after Main) : error up to about zrVel x 2 cycles + the input filter *)
				gZRef.Output.MeasuredZ := gAxis[AX_Z].Output.State.Position;
				stepTimer(IN := FALSE);
				fbZrMove[2].Execute := FALSE;
				fbZrHalt[2].Execute := TRUE;
				commandStep := 50;
			ELSIF fbZrMove[2].Done THEN
				(* MaxZ reached without a signal (no sensor, sensor not wired) *)
				stepTimer(IN := FALSE);
				fbZrMove[2].Execute := FALSE;
				zrFail := 3;
				commandStep := 60;
			ELSIF fbZrMove[2].Error OR fbZrMove[2].CommandAborted THEN
				zrFail := 4;
				commandStep := 190;
			ELSIF stepTimer.Q THEN
				zrFail := 6;
				commandStep := 190;
			END_IF

		50: (* braking on the sensor *)
			stepTimer(IN := TRUE, PT := T#5s);

			IF fbZrHalt[2].Done THEN
				stepTimer(IN := FALSE);
				fbZrHalt[2].Execute := FALSE;
				commandStep := 60;
			ELSIF fbZrHalt[2].Error OR fbZrHalt[2].CommandAborted THEN
				zrFail := 4;
				commandStep := 190;
			ELSIF stepTimer.Q THEN
				zrFail := 6;
				commandStep := 190;
			END_IF

		60: (* Z back up to SafeZ - also after ErrorId 2 / 3 *)
			fbZrMove[2].Position := gZRef.Input.SafeZ;
			fbZrMove[2].Velocity := zrMoveVel;
			fbZrMove[2].Execute := TRUE;
			stepTimer(IN := FALSE);
			commandStep := 61;

		61:
			stepTimer(IN := TRUE, PT := T#60s);

			IF fbZrMove[2].Done THEN
				stepTimer(IN := FALSE);
				fbZrMove[2].Execute := FALSE;
				zrActive := FALSE;
				IF zrFail = 0 THEN
					gZRef.Output.Head := gZRef.Input.Head;
					gZRef.Output.Done := TRUE;
					commandStep := 100;
				ELSE
					gZRef.Output.ErrorId := zrFail;
					commandStep := 200;
				END_IF
			ELSIF fbZrMove[2].Error OR fbZrMove[2].CommandAborted THEN
				zrFail := 4;
				commandStep := 190;
			ELSIF stepTimer.Q THEN
				zrFail := 6;
				commandStep := 190;
			END_IF

		190: (* a move failed : brake what this cycle still moves, no result *)
			stepTimer(IN := FALSE);
			FOR i := 0 TO 2 DO
				IF fbZrMove[i].Busy THEN
					fbZrHalt[i].Execute := TRUE;
				END_IF
				fbZrMove[i].Execute := FALSE;
			END_FOR
			gZRef.Output.ErrorId := zrFail;
			zrActive := FALSE;
			commandStep := 200;

		100:
			zrActive := FALSE;(* Complete - gZRef.Output.MeasuredZ / Head *)

		200:
			zrActive := FALSE;(* failed - gZRef.Output.ErrorId *)
	END_CASE

END_ACTION

ACTION act_ZRef:
	(* every cycle : input check for the next command, end of a measurement that was left (STOP, ABORT, E-stop, handwheel),
	   release of the halts, status *)
	act_ZRefCheck;

	IF zrActive AND (cncCommand <> E_ACT_MEASURE_Z OR DI_MPG_Jog_Enable OR emergencyLatched) THEN
		(* brake what the measurement still moves, the result is not valid *)
		FOR i := 0 TO 2 DO
			IF fbZrMove[i].Busy THEN
				fbZrHalt[i].Execute := TRUE;
			END_IF
			fbZrMove[i].Execute := FALSE;
		END_FOR
		gZRef.Output.ErrorId := 5;
		zrActive := FALSE;
		IF cncCommand = E_ACT_MEASURE_Z THEN
			commandStep := 200; (* handwheel : the command ends *)
		END_IF
	END_IF

	IF NOT zrActive THEN
		FOR i := 0 TO 2 DO
			IF fbZrHalt[i].Done OR fbZrHalt[i].Error OR fbZrHalt[i].CommandAborted THEN
				fbZrHalt[i].Execute := FALSE;
			END_IF
		END_FOR
	END_IF

	gZRef.Output.Sensor := DI_ZRef_Sensor;
	gZRef.Output.Busy := zrActive;
	IF zrActive THEN
		gZRef.Output.Step := commandStep;
	ELSE
		gZRef.Output.Step := 0;
	END_IF

END_ACTION
```

#### Action_WorkOffset.st - Work offset actions
```iecst
ACTION act_WorkOffset:
	(* Work offsets G54..G57 (HMI work offset card) : machine position of the program origin per offset. Apply (HMI) takes the
	   table and the active offset over while the CNC is idle (refused otherwise : Output.Rejected). act_Start /
	   act_MoveBlock set the active offset as the standard frame SCS1 (MC_BR_SetStandardFrame, translation only) right before
	   the run, so program and MDI coordinates are relative to that origin : machine = program + offset.
	   While the active offset and the frame set last are both 0 (the default) nothing is set
	   (program coordinates = machine coordinates). Single-axis moves (jog, ManualMove, teach positions), homing, the ring
	   buffer stay in machine coordinates.
	   In-program G54..G59 select the frame table frame (SCS3) of mapp Motion, which is not configured - not used here *)

	(* Apply : only while idle and with sane values - a run in progress keeps its frame *)
	IF gWorkOffset.Input.Command.Apply THEN
		gWorkOffset.Input.Command.Apply := FALSE;
		woOk := cncCommand = E_ACT_IDLE AND NOT programAlive AND woStep = 0
			AND gWorkOffset.Input.Parameter.Active <= 3;
		FOR woIdx := 0 TO 3 DO
			woOk := woOk AND ABS(gWorkOffset.Input.Parameter.Offset[woIdx].X) <= C_WO_MAX
				AND ABS(gWorkOffset.Input.Parameter.Offset[woIdx].Y) <= C_WO_MAX
				AND ABS(gWorkOffset.Input.Parameter.Offset[woIdx].Z) <= C_WO_MAX;
		END_FOR
		IF woOk THEN
			FOR woIdx := 0 TO 3 DO
				gWorkOffset.Output.Offset[woIdx] := gWorkOffset.Input.Parameter.Offset[woIdx];
			END_FOR
			gWorkOffset.Output.Active := gWorkOffset.Input.Parameter.Active;
		END_IF
		gWorkOffset.Output.Rejected := NOT woOk;
	END_IF

	(* frame of the active offset (translation only) *)
	IF gWorkOffset.Output.Active <= 3 THEN
		woIdx := gWorkOffset.Output.Active;
	ELSE
		woIdx := 0;
	END_IF
	woWant.Pos.X := gWorkOffset.Output.Offset[woIdx].X;
	woWant.Pos.Y := gWorkOffset.Output.Offset[woIdx].Y;
	woWant.Pos.Z := gWorkOffset.Output.Offset[woIdx].Z;

	(* set before a run only when an offset is or was in use - it is set again before every run, so a frame that mapp
	   Motion resets at the end of a program (modal data) is back for the next one *)
	woNeed := woWant.Pos.X <> 0.0 OR woWant.Pos.Y <> 0.0 OR woWant.Pos.Z <> 0.0
		OR woSet.Pos.X <> 0.0 OR woSet.Pos.Y <> 0.0 OR woSet.Pos.Z <> 0.0;
	gWorkOffset.Output.InUse := woNeed;

	(* the run that requested the frame is over (also STOP / ABORT while it was set) *)
	IF (woStep = 100 OR woStep = 200) AND cncCommand = E_ACT_IDLE THEN
		woStep := 0;
	END_IF

	CASE woStep OF
		1: (* requested by act_Start / act_MoveBlock *)
			woTimer(IN := FALSE);
			gWorkOffset.Output.Error := FALSE;
			gWorkOffset.Output.ErrorID := 0;
			fbWorkFrame.Frame := woWant;
			fbWorkFrame.Execute := TRUE;
			woStep := 10;

		10:
			woTimer(IN := TRUE, PT := T#2s);

			IF fbWorkFrame.Done THEN
				woTimer(IN := FALSE);
				fbWorkFrame.Execute := FALSE;
				woSet := fbWorkFrame.Frame;
				woStep := 100;
			ELSIF fbWorkFrame.Error OR woTimer.Q THEN
				(* the run is not started : it would run at the wrong place *)
				woTimer(IN := FALSE);
				fbWorkFrame.Execute := FALSE;
				gWorkOffset.Output.Error := TRUE;
				gWorkOffset.Output.ErrorID := fbWorkFrame.ErrorID;
				woStep := 200;
			END_IF

		100:
			;(* set - the action goes on with the run *)

		200:
			;(* failed - the action ends with 200 *)
	END_CASE

END_ACTION
```

#### Action_HeadOffset.st - Head offset actions
```iecst
ACTION act_HeadOffset:
	(* Head (tool) offsets : the axis positions refer to the reference head tip, each head's working point sits at its offset
	   from there (HMI head table, H1..H4 = PlcId). Only one head is mounted at a time (HMI plugin structure), so the offset of
	   the mounted head (ActiveHead) holds for every run. Apply (HMI) takes the table and the mounted head over while the CNC is
	   idle (refused otherwise : Output.Rejected). act_Start / act_MoveBlock set minus that offset as the standard
	   frame SCS2 (MC_BR_SetStandardFrame, translation only) right before the run, so the head's working point follows the
	   program : machine = program - offset.
	   While the mounted head's offset and the frame set last are both 0 (the default, ActiveHead 0 or the reference head)
	   nothing is set. Single-axis moves (jog, ManualMove, teach positions), homing, the ring
	   buffer stay at the reference head tip.
	   mapp tool tables (MC_BR_SetToolTable / MC_BR_SetToolPar) are not used : the axes group has no tool feature configured *)

	(* Apply : only while idle and with sane values - a run in progress keeps its frame *)
	IF gHeadOffset.Input.Command.Apply THEN
		gHeadOffset.Input.Command.Apply := FALSE;
		hoOk := cncCommand = E_ACT_IDLE AND NOT programAlive AND hoStep = 0
			AND gHeadOffset.Input.Parameter.ActiveHead <= 4;
		FOR hoIdx := 1 TO 4 DO
			hoOk := hoOk AND ABS(gHeadOffset.Input.Parameter.Offset[hoIdx].X) <= C_HO_MAX
				AND ABS(gHeadOffset.Input.Parameter.Offset[hoIdx].Y) <= C_HO_MAX
				AND ABS(gHeadOffset.Input.Parameter.Offset[hoIdx].Z) <= C_HO_MAX;
		END_FOR
		IF hoOk THEN
			FOR hoIdx := 1 TO 4 DO
				gHeadOffset.Output.Offset[hoIdx] := gHeadOffset.Input.Parameter.Offset[hoIdx];
			END_FOR
			gHeadOffset.Output.ActiveHead := gHeadOffset.Input.Parameter.ActiveHead;
		END_IF
		gHeadOffset.Output.Rejected := NOT hoOk;
	END_IF

	(* frame of the mounted head : minus its offset (translation only), none = 0 *)
	hoWant.Pos.X := 0.0;
	hoWant.Pos.Y := 0.0;
	hoWant.Pos.Z := 0.0;
	IF gHeadOffset.Output.ActiveHead >= 1 AND gHeadOffset.Output.ActiveHead <= 4 THEN
		hoIdx := gHeadOffset.Output.ActiveHead;
		hoWant.Pos.X := -gHeadOffset.Output.Offset[hoIdx].X;
		hoWant.Pos.Y := -gHeadOffset.Output.Offset[hoIdx].Y;
		hoWant.Pos.Z := -gHeadOffset.Output.Offset[hoIdx].Z;
	END_IF

	(* set before a run only when an offset is or was in use - it is set again before every run, so a frame that mapp
	   Motion resets at the end of a program (modal data) is back for the next one *)
	hoNeed := hoWant.Pos.X <> 0.0 OR hoWant.Pos.Y <> 0.0 OR hoWant.Pos.Z <> 0.0
		OR hoSet.Pos.X <> 0.0 OR hoSet.Pos.Y <> 0.0 OR hoSet.Pos.Z <> 0.0;
	gHeadOffset.Output.InUse := hoNeed;

	(* the run that requested the frame is over (also STOP / ABORT while it was set) *)
	IF (hoStep = 100 OR hoStep = 200) AND cncCommand = E_ACT_IDLE THEN
		hoStep := 0;
	END_IF

	CASE hoStep OF
		1: (* requested by act_Start / act_MoveBlock *)
			hoTimer(IN := FALSE);
			gHeadOffset.Output.Error := FALSE;
			gHeadOffset.Output.ErrorID := 0;
			fbHeadFrame.Frame := hoWant;
			fbHeadFrame.Execute := TRUE;
			hoStep := 10;

		10:
			hoTimer(IN := TRUE, PT := T#2s);

			IF fbHeadFrame.Done THEN
				hoTimer(IN := FALSE);
				fbHeadFrame.Execute := FALSE;
				hoSet := fbHeadFrame.Frame;
				hoStep := 100;
			ELSIF fbHeadFrame.Error OR hoTimer.Q THEN
				(* the run is not started : the head would work at the wrong place *)
				hoTimer(IN := FALSE);
				fbHeadFrame.Execute := FALSE;
				gHeadOffset.Output.Error := TRUE;
				gHeadOffset.Output.ErrorID := fbHeadFrame.ErrorID;
				hoStep := 200;
			END_IF

		100:
			;(* set - the action goes on with the run *)

		200:
			;(* failed - the action ends with 200 *)
	END_CASE

END_ACTION
```

#### Variables.var - Local variables
```iecst
VAR
	fbCnc : MpCnc3Axis;
	CncParameters : MpCnc3AxisParType;
	bootPowerDone : BOOL := FALSE; (*servo powered once after boot*)
	initThenHome : BOOL := FALSE; (*INIT continues with HOME (HMI) or stops after power on (boot)*)
	cmdAllowed : BOOL := FALSE; (*preconditions of the command in the mailbox*)
END_VAR
(*Emergency stop*)
VAR
	emergencyLatched : BOOL := FALSE; (*set by the E-stop button, cleared by RESET once released*)
	emergencyTimer : TON; (*power off at the latest after this, even if the axes have not stopped*)
END_VAR
(*Main*)
VAR
	i : USINT := 0;
	cncCommand : E_CNC_ACTION := E_ACT_IDLE;
	commandStep : USINT := 0;
	stepTimer : TON;
END_VAR
(*Axis Reset*)
VAR
	fbAxisReset : ARRAY[0..2] OF MC_Reset;
END_VAR
(*X Axis Deviation Compensation - mapp Motion*)
VAR
	fbMechDevCompX : MC_BR_MechDeviationComp;
END_VAR
(*M Function - mapp Motion*)
VAR
	fbMFunction : ARRAY[0..7] OF MC_BR_MFunction; (*0 = M41, 1 = M42, 2 = M44, 3 = M45, 4 = M61, 5 = M62 (async), 6 = M50, 7 = M51 (blocking, no function - reset at once by act_MSpare)*)
	fbMFunctionSpare : ARRAY[0..7] OF MC_BR_MFunction; (*0..7 = M52..M59 : rest of the blocking range 50..59 (Config_6) - no function on this machine, reset at once by act_MSpare so a program does not wait there for ever*)
	mfSpareLast : USINT := 0; (*last of M50..M59 passed since power-up, 0 = none - diagnosis only*)
	mfClear : BOOL := FALSE; (*no program / E-stop : discharge and laser off, M41 / M61 held in reset*)
	programStarted : BOOL := FALSE; (*a production run was started by START (not MDI)*)
	programAlive : BOOL := FALSE; (*a program runs or is paused (HALT, single step, M01) : fbCnc.MoveActive OR programHeld*)
	programEndTrig : F_TRIG; (*end of programAlive*)
END_VAR
(*Single step / optional stop (M01) - gCncRun*)
VAR
	fbOptStop : MC_BR_OptionalStop; (*the program stops at M01 while gCncRun.Input.OptionalStop is set*)
	programHeld : BOOL := FALSE; (*the program waits for CONTINUE : interrupted (HALT, single step), standing at M01 or waiting before its real run (start at line)*)
	stepHold : BOOL := FALSE; (*the program stopped by itself (single step, M01, start at line waiting) : act_Start hands over to the mailbox like after HALT, so CONTINUE is taken*)
END_VAR
(*Start at line (E_ACT_START_AT_LINE) - gCncRun*)
VAR
	lineStartRun : BOOL := FALSE; (*the alive program was started by E_ACT_START_AT_LINE*)
	lineStartPrep : BOOL := FALSE; (*that program is before its real run : simulation up to the start line, repositioning, waiting*)
	lineStartWait : BOOL := FALSE; (*that program waits for CONTINUE before or after the repositioning*)
END_VAR
(*MDI (act_MoveBlock)*)
VAR
	mdiDoneOld : BOOL := FALSE; (*MoveDone was already set when the block was given : not this block's until it falls*)
	mdiAbortOld : BOOL := FALSE; (*the same for CommandAborted*)
END_VAR
(*Heads - only the active head (gActiveHead) is taken (Action_Head.st)*)
VAR
	headDispOk : BOOL := TRUE; (*the dispenser may be switched on : gActiveHead is 0 (not known) or the dispenser*)
	headLaserOk : BOOL := TRUE; (*the laser may be switched on : gActiveHead is 0 (not known) or the laser*)
	headRefuse : USINT := 0; (*head refused in this cycle (HEAD_ constants), 0 = none*)
	headMfTrig : ARRAY[0..5] OF R_TRIG; (*rising edge of fbMFunction[0..5].Value*)
	headRunTrig : R_TRIG; (*a run starts (programAlive) : the last refusal is cleared*)
END_VAR
(*Teach positions*)
VAR
	teachSum : LREAL := 0.0; (*only references C_TP1_1 .. C_TP4_3 in _INIT so that the global PVs are created on the target*)
END_VAR
(*Z reference measurement (Action_ZRef.st) - single-axis moves of its own, machine coordinates*)
VAR
	fbZrMove : ARRAY[0..2] OF MC_MoveAbsolute; (*0 = X, 1 = Y, 2 = Z - only used by the measurement*)
	fbZrHalt : ARRAY[0..2] OF MC_Halt;
	zrActive : BOOL := FALSE; (*measurement running (cncCommand = E_ACT_MEASURE_Z, steps 10..61)*)
	zrFail : USINT := 0; (*ErrorId to report once Z is back at SafeZ*)
	zrVel : REAL := 0.0; (*search velocity [mm/s]*)
	zrMoveVel : REAL := 0.0; (*velocity of the other moves = SystemSpeed, like ManualMove [mm/s]*)
END_VAR
(*Work offsets G54..G57 (Action_WorkOffset.st) - the active offset is set as the standard frame SCS1 before a run*)
VAR
	fbWorkFrame : MC_BR_SetStandardFrame;
	woStep : USINT := 0; (*frame engine: 0 idle, 1 requested by act_Start / act_MoveBlock, 10 setting, 100 set, 200 failed*)
	woNeed : BOOL := FALSE; (*the frame has to be set before a run : the active offset or the frame set last is not 0*)
	woWant : McFrameType; (*frame of the active offset*)
	woSet : McFrameType; (*frame set last since boot (the axes group starts with 0)*)
	woOk : BOOL := FALSE; (*Apply accepted*)
	woIdx : USINT := 0;
	woTimer : TON;
END_VAR
(*Head (tool) offsets (Action_HeadOffset.st) - minus the mounted head's offset is set as the standard frame SCS2 before a run*)
VAR
	fbHeadFrame : MC_BR_SetStandardFrame;
	hoStep : USINT := 0; (*frame engine: 0 idle, 1 requested by act_Start / act_MoveBlock, 10 setting, 100 set, 200 failed*)
	hoNeed : BOOL := FALSE; (*the frame has to be set before a run : the active head's offset or the frame set last is not 0*)
	hoWant : McFrameType; (*frame of the mounted head (minus its offset)*)
	hoSet : McFrameType; (*frame set last since boot (the axes group starts with 0)*)
	hoOk : BOOL := FALSE; (*Apply accepted*)
	hoIdx : USINT := 0;
	hoTimer : TON;
END_VAR
VAR CONSTANT
	C_ZREF_PROBE_VEL : REAL := 2.0; (*default search velocity of the Z reference measurement [mm/s]*)
	C_ZREF_MAX_VEL : REAL := 10.0; (*largest search velocity accepted [mm/s]*)
	C_ZREF_MOVE_VEL : REAL := 50.0; (*velocity of the other measurement moves when SystemSpeed is 0 [mm/s]*)
	C_ZREF_MAX_SEARCH : LREAL := 50.0; (*largest search range MaxZ - StartZ [mm]*)
	C_ZREF_ACC : REAL := 500.0; (*acceleration / deceleration of the measurement moves and halts [mm/s2] - as AxisManual DEFAULT_ACC / DEFAULT_DEC*)
	C_WO_MAX : LREAL := 10000.0; (*largest work offset accepted by Apply [mm]*)
	C_HO_MAX : LREAL := 1000.0; (*largest head offset accepted by Apply [mm]*)
END_VAR
```

### Program Logical/Cnc/OpMode (IEC) - Operating mode (auto / manual) and handwheel selection

#### Cyclic.st - Cyclic code
```iecst
PROGRAM _CYCLIC

	(* mode selector switch not wired : HMI selects the mode. A change is taken over only while the CNC is idle *)
	IF gEquipment.Output.Status.CurrentAction = E_ACT_IDLE AND NOT gEquipment.Output.Status.ProgramActive AND NOT gEquipment.Output.State.Move THEN
		DI_Auto := NOT gEquipment.Input.Command.ManualMode;
	END_IF

	Action_ControlButton;

	(* MPG has no enable switch : an axis selected on the MPG means MPG mode (blocks AxisManual) *)
	DI_MPG_Jog_Enable := DI_MPG_AxisX OR DI_MPG_AxisY OR DI_MPG_AxisZ;

END_PROGRAM
```

#### Init.st - Init code
```iecst
PROGRAM _INIT

END_PROGRAM
```

#### Exit.st - Exit code
```iecst
PROGRAM _EXIT
END_PROGRAM
```

#### Variables.var - Local variables
```iecst
VAR
	ManualModeTrigger : F_TRIG := (0);
END_VAR
```

#### Action_ControlButton.st
```iecst
ACTION Action_ControlButton:

	(* auto -> manual : stop CNC and discharge *)
	ManualModeTrigger(CLK := DI_Auto);

	IF ManualModeTrigger.Q THEN
		gDispenser.Input.Command.Discharge := FALSE;
		gEquipment.Input.CncCommand := E_ACT_STOP;
	END_IF

END_ACTION
```

### Program Logical/Cnc/PrgShare (IEC) - Network share of the CNC programs (file device CNC_PrgDir)

#### Cyclic.st - Cyclic code
```iecst
PROGRAM _CYCLIC

	CASE step OF
		0: (* link the network share as the file device of the CNC programs *)
			fbDevLink.enable := TRUE;
			fbDevLink.pDevice := ADR(deviceName);
			fbDevLink.pParam := ADR(shareParam);
			fbDevLink();

			IF fbDevLink.status = ERR_OK THEN
				linked := TRUE;
				linkStatus := 0;
				step := 10;
			ELSIF fbDevLink.status <> ERR_FUB_BUSY AND fbDevLink.status <> ERR_FUB_ENABLE_FALSE THEN
				linkStatus := fbDevLink.status;
				sysError := FileIoGetSysError();
				fbDevLink.enable := FALSE;
				fbDevLink();
				step := 20;
			END_IF

		10: (* linked *)

		20: (* failed : try again after 10 s (share or PC not reachable yet) *)
			retryTimer(IN := TRUE, PT := T#10s);
			IF retryTimer.Q THEN
				retryTimer(IN := FALSE);
				step := 0;
			END_IF

	END_CASE

END_PROGRAM
```

#### Init.st - Init code
```iecst
PROGRAM _INIT
END_PROGRAM
```

#### Exit.st - Exit code
```iecst
PROGRAM _EXIT
END_PROGRAM
```
